RoboDK station: robotic_car_painting_cell.rdk

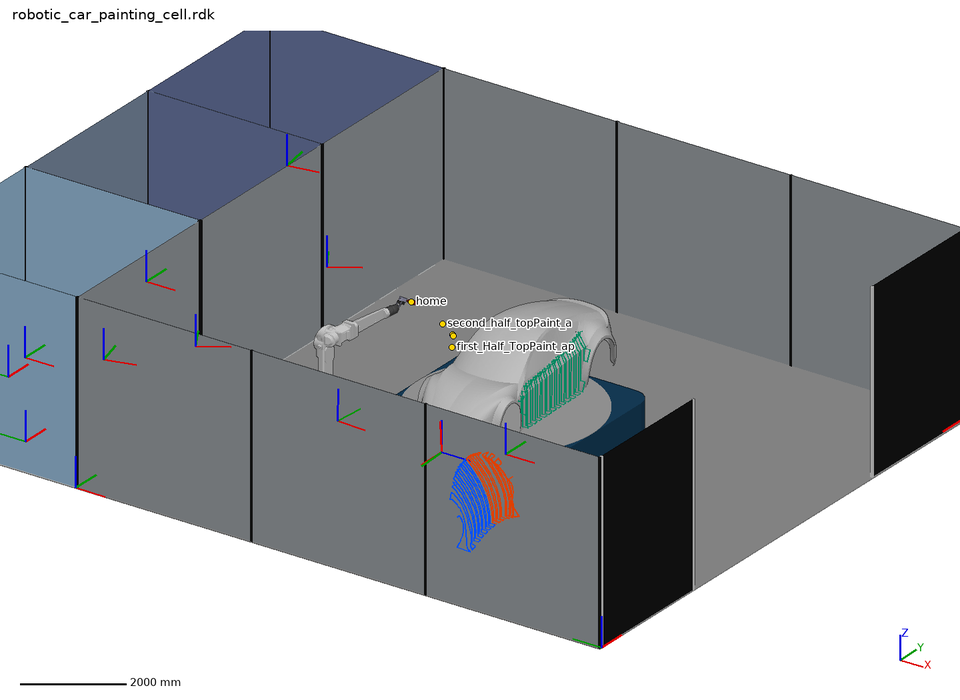
[picture v0: the station drawn from its stored meshes, robots at their saved joint values, targets as dots, program paths as lines]
Station robotic_car_painting_cell (saved by RoboDK 6.1.1). Poses are relative to the parent item; angles as X-Y-Z fixed-axis rotations.
  - frame ABB IRB 5500-27 Base at (-2375.69, -2107.7, 876.55) mm, rotated rx -0.57 ry -0.3 rz -4.19 deg
    - robot ABB IRB 5500-27: 6 axes, payload 16 kg, reach 2200 mm, repeatability 0.15 mm, weight 600 kg
        modified DH rows (alpha deg, a mm, theta deg, d mm): 0, 0, 0, 436; -90, 0, -90, -5; 0, 1300, 0, 0; -90, 0, -90, 1510.5; 35, 0, 0, 79.169; -70, 0, 180, 79.169
        base shift (0, 0, 0) mm, rotated rx 0 ry 0 rz 90 deg
        joint limits [-104, -65, -70, -719, -719, -720] to [104, 150, 70, 719, 719, 720]; home [0, 0, 0, 0, 0, 0]; saved at [0, 0, 0, 0, 0, 0]
      - tool Paint gun, TCP at (50, 0, 450) mm, rotated rx 0 ry 30 rz 0 deg, size 203.2 x 279.7 x 471.5 mm
    - target home (joint target) at (5, 2172.1, 1686) mm, rotated rx 180 ry 60 rz -90 deg; joints [0, 0, 0, 0, 0, 0, 0] of ABB IRB 5500-27
    - target first_Half_TopPaint_app (joint target) at (1861.11, 1119.96, 1686) mm, rotated rx 180 ry 60 rz -148.83 deg; joints [-58.83, 0, 0, 0, 0, 0, -69.91] of ABB IRB 5500-27
    - target second_half_topPaint_app (joint target) at (1072.69, 1796.81, 1679.78) mm, rotated rx 180 ry 59.9 rz -120.7 deg; joints [-30.7, -3.5, 3.6, 0, 0, 0, -28] of ABB IRB 5500-27
    - target second_to_home (joint target) at (1519.79, 1551.86, 1686) mm, rotated rx 180 ry 60 rz -134.27 deg; joints [-44.27, 0, 0, 0, 0, 0, -33.04] of ABB IRB 5500-27
    - target sidePaintApp (joint target) at (1560.69, 1510.73, 1686) mm, rotated rx 180 ry 60 rz -135.8 deg; joints [-45.8, 0, 0, 0, 0, 0, -170] of ABB IRB 5500-27
  - frame Turntable 1 Base at (0, 0, 0) mm
    - robot Turntable 1: 1 axes
        modified DH rows (alpha deg, a mm, theta deg, d mm): 0, 0, 0, 0
        base shift (0, 0, 1000) mm
        joint limits [-1000] to [1000]; home [0]; saved at [0]
      - frame carFrame at (0, -2099.21, -116.89) mm, rotated rx 90 ry 0 rz 0 deg
        - object carBodyTesla at (0, 0, 0) mm, size 1894.9 x 1628.8 x 4824.9 mm, geometry from carBodyTesla.STEP
        - frame FrameSidePaint at (0, 0, 0) mm, rotated rx -92.52 ry -89.99 rz 2.4 deg
          - object carSidePaint at (0, 0, 0) mm, geometry from       
        - frame FrameTopPaint at (0, 0, 0) mm, rotated rx 90 ry -3.48 rz 90 deg
          - object carTopPaint at (0, 0, 0) mm, rotated rx 90 ry 0 rz 86.52 deg, geometry from pacity
  - machining project first_half_topPaint: rotZ(0) | rotX(0)*rotY(0) | onStart | onPathStart | onApproach | onPoint | onRetract | onFinish | SetRPM(%1) | SetTool(%1) | Extruder(%1) | default | default | OutOnMov(%1) | OutOffMov(%1) | onPathFinish | M_RunCode(%1)
  - program first_half_topPaint (530 instructions, listed below)
  - machining project Path2 settings: rotZ(0) | rotX(0)*rotY(0) | rotz(0) | onStart | onPathStart | onApproach | onPoint | onRetract | onFinish | SetRPM(%1) | SetTool(%1) | Extruder(%1) | default | default | OutOnMov(%1) | OutOffMov(%1) | onPathFinish | M_RunCode(%1)
  - program second_half_topPaint (492 instructions, listed below)
  - machining project Path3 settings: rotZ(0) | rotX(0)*rotY(0) | rotz(90) | onStart | onPathStart | onApproach | onPoint | onRetract | onFinish | SetRPM(%1) | SetTool(%1) | Extruder(%1) | default | default | OutOnMov(%1) | OutOffMov(%1) | onPathFinish | M_RunCode(%1)
  - program side_paint (1096 instructions, listed below)
  - program second_half_topPaint_startP (3 instructions, listed below)
  - program first_half_topPaint_startP (3 instructions, listed below)
  - program second_to_First_conn (3 instructions, listed below)
  - program CarTopPaintMain (3 instructions, listed below)
  - program sidePaint_startP (3 instructions, listed below)
  - program CarSidePaintMain (1 instructions, listed below)
  - program Home (3 instructions, listed below)
  - object robot_stand at (-2371.87, -2116.55, 0) mm, size 1000 x 999.7 x 874.6 mm
  - frame Components at (-5797.63, -5825.6, 0) mm
    - frame Fence 1 Frame at (0, 0, 0) mm
      - object Fence 1 at (0, 0, 0) mm, size 12050 x 12050 x 4010 mm
    - frame Fence 1 Frame at (-4009.44, 0, 0) mm
      - object Fence 1 at (0, 0, 0) mm, size 4050 x 4050 x 4010 mm
    - frame Fence 1 Frame at (-3997.18, 4026.78, 0) mm
      - object Fence 1 at (0, 0, 0) mm, size 4050 x 4050 x 4010 mm
    - frame Fence 1 Frame at (-3995.72, 8010.06, 0) mm
      - object Fence 1 at (0, 0, 0) mm, size 4050 x 4050 x 4010 mm
    - frame Fence 1 Frame at (11995.78, 12001.82, 0) mm, rotated rx 0 ry 0 rz -90.05 deg
      - object Fence 1 at (0, 0, 0) mm, size 3050 x 50 x 4000 mm
    - frame Fence 2 Frame at (12049.84, 56.15, 0) mm, rotated rx 0 ry 0 rz 89.84 deg
      - object Fence 2 at (0, 0, 0) mm, size 3050 x 50 x 4000 mm
    - frame Box 1 Frame at (-1567.64, 10491.56, 0) mm, rotated rx 0 ry 0 rz 32.89 deg
      - object Box 1 at (0, 0, 0) mm, size 1000 x 1000 x 500 mm, geometry from cube.sld
    - frame Sphere 1 Frame at (-2358.15, 10303.8, 1975.89) mm, rotated rx 0 ry 0 rz 9.39 deg
      - object Sphere 1 at (0, -1304.1, -1382.72) mm, size 1000 x 1000 x 1000 mm, geometry from sph.sld
    - frame Prism 2 Frame at (-2731.49, 4804.46, 0) mm, rotated rx 0 ry 0 rz 14.89 deg
      - object Prism 2 at (0, 0, 0) mm, size 1000 x 1000 x 500 mm, geometry from prism.sld
    - frame Table 1 Frame at (-1857.36, 1009.43, 39.55) mm, rotated rx 0 ry 0 rz 90.42 deg
      - frame Table 1 Plane Frame at (-585.26, 0, 1600) mm
      - object Table 1 at (0, 0, 0) mm, size 2000 x 1000 x 1600 mm
    - frame Cone 1 Frame at (-1643.96, 6288.26, 0) mm, rotated rx 0 ry 0 rz 30.73 deg
      - object Cone 1 at (0, 0, 0) mm, size 700 x 700 x 600 mm
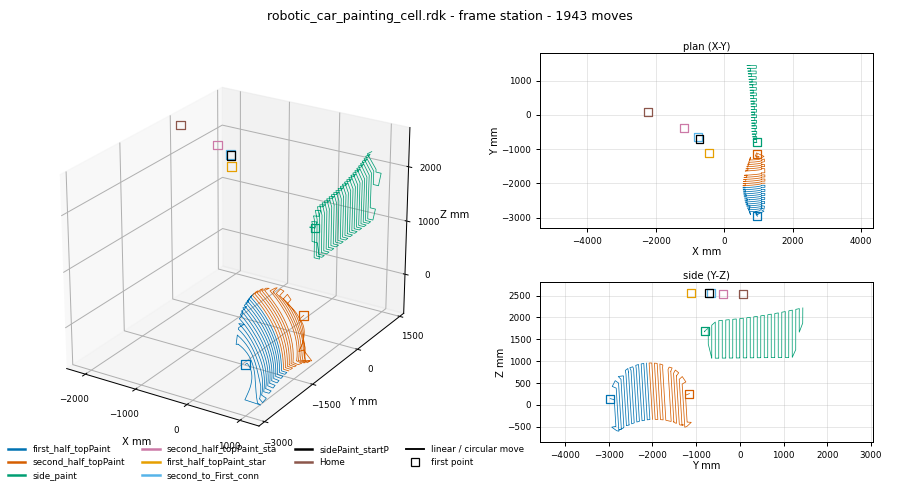
[picture p0: tool path of robotic_car_painting_cell.rdk in frame station, 1943 of 1943 moves have a stored position in this frame; points joined in program order, loops and branches not executed]

--- program first_half_topPaint (robot ABB IRB 5500-27) ---
  Smooth(1)
  Set speed (1000.0 mm/s)
  Set Ref.: FrameTopPaint
  Set Tool: Paint gun
  Show Paint gun
  MoveJ 1 to (-684.51, 907.52, 971.03) mm, rotated rx 106.25 ry 20.82 rz -12.55 deg; joints [-74.794, -12.721, 37.414, 15.51, -31.42, 69.743, -69.91]
  MoveL 2 to (-684.51, 907.52, 971.03) mm, rotated rx 106.25 ry 20.82 rz -12.55 deg; joints [-74.794, -12.721, 37.414, 15.51, -31.42, 69.743, -69.91]
  MoveL 3 to (-715.08, 815.97, 944.87) mm, rotated rx 106.25 ry 20.82 rz -12.55 deg; joints [-70.189, -11.053, 37.131, 20.085, -29.663, 64.32, -69.91]
  MoveL 4 to (-715.08, 815.97, 944.87) mm, rotated rx 106.25 ry 20.82 rz -12.55 deg; joints [-70.189, -11.053, 37.131, 20.085, -29.663, 64.32, -69.91]
  Set speed (50.0 mm/s)
  MoveL 5 to (-727.69, 815.97, 958.3) mm, rotated rx 115.21 ry 38.9 rz -3.5 deg; joints [-72.492, -7.954, 36.366, 53.545, -66.561, 43.021, -69.91]
  MoveL 6 to (-741.38, 815.97, 970.44) mm, rotated rx 121.28 ry 37.31 rz -1.34 deg; joints [-71.643, -9.484, 34.92, 41.962, -56.112, 42.571, -69.91]
  MoveL 7 to (-756.1, 815.97, 981.34) mm, rotated rx 127.91 ry 34.94 rz 0.84 deg; joints [-70.269, -10.891, 33.104, 25.851, -42.702, 44.586, -69.91]
  MoveL 8 to (-771.81, 815.97, 991.01) mm, rotated rx 147.14 ry 44.4 rz 22.43 deg; joints [-72.285, -8.078, 30.032, 38.203, -68.24, 34.256, -69.91]
  MoveL 9 to (-788.18, 815.97, 999.35) mm, rotated rx 152.65 ry 38.6 rz 23.9 deg; joints [-70.353, -9.282, 27.683, 18.408, -52.224, 37.943, -69.91]
  MoveL 10 to (-804.72, 815.97, 1006.28) mm, rotated rx 157.1 ry 32.58 rz 24.14 deg; joints [-67.802, -9.883, 25.248, -7.481, -33.792, 47.461, -69.91]
  MoveL 11 to (-821.7, 815.97, 1012.06) mm, rotated rx 171.62 ry 31.52 rz 45.71 deg; joints [-69.524, -6.36, 20.448, 5.697, -60.164, 39.026, -69.91]
  MoveL 12 to (-839.09, 815.97, 1016.77) mm, rotated rx 172.06 ry 25.49 rz 43.55 deg; joints [-67.355, -6.129, 18.073, -13.153, -47.594, 47.333, -69.91]
  MoveL 13 to (-856.8, 815.97, 1020.47) mm, rotated rx 172.25 ry 20.32 rz 41.61 deg; joints [-65.459, -5.39, 15.854, -31.628, -37.033, 57.574, -69.91]
  MoveL 14 to (-879.91, 815.97, 1023.85) mm, rotated rx 172.07 ry 15.06 rz 39.99 deg; joints [-63.836, -3.875, 13.191, -50.671, -28.335, 70.216, -69.91]
  MoveL 15 to (-903.07, 815.97, 1025.78) mm, rotated rx 171.26 ry 11.43 rz 39.86 deg; joints [-63.298, -1.925, 10.503, -57.68, -27.796, 76.89, -69.91]
  MoveL 16 to (-926.28, 815.97, 1026.44) mm, rotated rx 169.77 ry 9.41 rz 41.6 deg; joints [-63.721, 0.361, 7.673, -51.962, -34.901, 76.409, -69.91]
  MoveL 17 to (-949.54, 815.97, 1025.94) mm, rotated rx 167.69 ry 9.08 rz 45.24 deg; joints [-64.892, 2.979, 4.812, -39.109, -46.426, 72.324, -69.91]
  MoveL 18 to (-972.84, 815.97, 1024.4) mm, rotated rx 162.64 ry 4.98 rz 31.07 deg; joints [-63.067, 2.797, 5.746, -87.371, -13.884, 106.328, -69.91]
  MoveL 19 to (-996.1, 815.97, 1021.9) mm, rotated rx 159.46 ry 7.32 rz 37.29 deg; joints [-65.349, 5.612, 2.717, -48.527, -38.544, 85.33, -69.91]
  MoveL 20 to (-1019.16, 815.97, 1018.56) mm, rotated rx 156.28 ry 11.18 rz 43.19 deg; joints [-67.612, 8.569, 0.499, -24.443, -55.69, 75.354, -69.91]
  MoveL 21 to (-1054.91, 815.97, 1011.84) mm, rotated rx 147.55 ry 8.73 rz 32.21 deg; joints [-67.708, 9.55, 0.627, -38.437, -41.429, 89.233, -69.91]
  MoveL 22 to (-1090.21, 815.97, 1003.5) mm, rotated rx 141.46 ry 15.3 rz 35.63 deg; joints [-70.243, 13.119, -0.752, -11.462, -57.847, 79.186, -69.91]
  MoveL 23 to (-1125.14, 815.97, 993.72) mm, rotated rx 135.68 ry 21.23 rz 35.98 deg; joints [-71.841, 16.239, -1.381, 6.343, -68.344, 74.883, -69.91]
  MoveL 24 to (-1159.69, 815.96, 982.62) mm, rotated rx 130.17 ry 26.09 rz 34.38 deg; joints [-72.775, 18.955, -1.682, 19.317, -75.346, 72.813, -69.91]
  MoveL 25 to (-1193.94, 815.97, 970.3) mm, rotated rx 120.68 ry 12.99 rz 20.14 deg; joints [-71.511, 17.84, -0.657, -10.346, -46.92, 91.196, -69.91]
  MoveL 26 to (-1227.25, 815.97, 957.05) mm, rotated rx 116.07 ry 14.96 rz 18.47 deg; joints [-71.999, 19.907, -0.984, -1.213, -50.466, 88.745, -69.91]
  MoveL 27 to (-1260.2, 815.97, 942.74) mm, rotated rx 112.21 ry 16.36 rz 16.46 deg; joints [-72.228, 21.731, -1.288, 5.505, -52.512, 87.03, -69.91]
  MoveL 28 to (-1293.17, 815.97, 928.47) mm, rotated rx 109.24 ry 17.29 rz 14.07 deg; joints [-72.243, 23.194, -1.506, 9.979, -52.843, 85.592, -69.91]
  MoveL 29 to (-1326.13, 815.97, 914.18) mm, rotated rx 106.48 ry 18.02 rz 12.4 deg; joints [-72.245, 24.912, -2.196, 14.357, -54.013, 84.608, -69.91]
  Set speed (1000.0 mm/s)
  MoveL 30 to (-1326.13, 815.97, 914.18) mm, rotated rx 106.48 ry 18.02 rz 12.4 deg; joints [-72.245, 24.912, -2.196, 14.357, -54.013, 84.608, -69.91]
  MoveL 31 to (-1338.15, 911.5, 941.16) mm, rotated rx 106.48 ry 18.02 rz 12.4 deg; joints [-74.918, 25.452, -3.974, 14.165, -56.682, 86.948, -69.91]
  Set speed (1000.0 mm/s)
  MoveL 32 to (-1426.8, 802.28, 1164.66) mm, rotated rx 159.74 ry 21.34 rz 28.53 deg; joints [-65.232, 18.141, -13.203, -64.298, -13.867, 90.288, -69.91]
  MoveL 33 to (-1440.26, 755.54, 1077.29) mm, rotated rx 159.74 ry 21.34 rz 28.53 deg; joints [-63.808, 19.217, -11.228, -70.076, -7.316, 90.993, -69.91]
  MoveL 34 to (-1440.26, 755.54, 1077.29) mm, rotated rx 159.74 ry 21.34 rz 28.53 deg; joints [-63.808, 19.217, -11.228, -70.076, -7.316, 90.993, -69.91]
  Set speed (50.0 mm/s)
  MoveL 35 to (-1392.1, 755.54, 1069.69) mm, rotated rx 159.42 ry 21.04 rz 29.31 deg; joints [-64.03, 17.502, -9.102, -59.847, -13.964, 85.038, -69.91]
  MoveL 36 to (-1343.82, 755.54, 1063.71) mm, rotated rx 159.05 ry 20.67 rz 30.24 deg; joints [-64.278, 15.856, -7.078, -52.603, -19.082, 81.124, -69.91]
  MoveL 37 to (-1295.44, 755.54, 1059.53) mm, rotated rx 158.62 ry 20.22 rz 31.39 deg; joints [-64.567, 14.305, -5.248, -46.409, -23.965, 78.169, -69.91]
  MoveL 38 to (-1246.95, 755.54, 1056.8) mm, rotated rx 158.2 ry 19.77 rz 32.55 deg; joints [-64.842, 12.754, -3.469, -41.574, -28.141, 76.122, -69.91]
  MoveL 39 to (-1198.41, 755.54, 1054.98) mm, rotated rx 157.76 ry 19.27 rz 33.81 deg; joints [-65.127, 11.251, -1.802, -37.325, -32.182, 74.6, -69.91]
  MoveL 40 to (-1154.25, 755.54, 1053.79) mm, rotated rx 157.34 ry 18.77 rz 35.08 deg; joints [-65.394, 9.936, -0.387, -33.798, -35.852, 73.57, -69.91]
  MoveL 41 to (-1110.09, 755.54, 1052.74) mm, rotated rx 156.9 ry 18.21 rz 36.48 deg; joints [-65.67, 8.687, 0.922, -30.459, -39.626, 72.814, -69.91]
  MoveL 42 to (-1065.93, 755.54, 1051.53) mm, rotated rx 156.43 ry 17.58 rz 38.07 deg; joints [-65.958, 7.531, 2.102, -27.18, -43.642, 72.297, -69.91]
  MoveL 43 to (-1021.8, 755.54, 1049.88) mm, rotated rx 157.68 ry 19.17 rz 34.06 deg; joints [-65.149, 3.751, 6.657, -35.423, -33.05, 72.924, -69.91]
  MoveL 44 to (-977.72, 755.54, 1047.5) mm, rotated rx 167.62 ry 20.43 rz 49.37 deg; joints [-66.013, 3.469, 6.21, -13.59, -56.701, 56.758, -69.91]
  MoveL 45 to (-933.75, 755.54, 1044.07) mm, rotated rx 170.23 ry 16.63 rz 43.58 deg; joints [-63.285, -0.433, 9.362, -37.882, -37.374, 65.285, -69.91]
  MoveL 46 to (-889.98, 755.54, 1039.27) mm, rotated rx 173.11 ry 14.65 rz 38.16 deg; joints [-60.377, -4.093, 13.488, -83.022, -6.548, 88.314, -69.91]
  MoveL 47 to (-860.05, 755.54, 1035) mm, rotated rx -179.66 ry 15.22 rz 55.82 deg; joints [-62.992, -3.267, 11.61, -25.717, -52.157, 51.737, -69.91]
  MoveL 48 to (-830.27, 755.54, 1029.79) mm, rotated rx -177.87 ry 15.22 rz 53.67 deg; joints [-61.924, -5.683, 14.166, -32.954, -44.629, 52.598, -69.91]
  MoveL 49 to (-800.66, 755.54, 1023.53) mm, rotated rx -176.11 ry 16.07 rz 52.51 deg; joints [-61.237, -7.933, 16.745, -36.847, -39.487, 51.96, -69.91]
  MoveL 50 to (-771.23, 755.54, 1016.08) mm, rotated rx -174.42 ry 17.74 rz 52.38 deg; joints [-61.049, -10.014, 19.323, -35.956, -37.616, 48.908, -69.91]
  MoveL 51 to (-746.52, 755.54, 1008.72) mm, rotated rx -173.04 ry 19.78 rz 53.06 deg; joints [-61.359, -11.624, 21.506, -30.839, -39.113, 44.159, -69.91]
  MoveL 52 to (-722.23, 755.54, 1000.38) mm, rotated rx -171.69 ry 22.36 rz 54.42 deg; joints [-62.128, -13.046, 23.699, -22.211, -43.408, 37.945, -69.91]
  MoveL 53 to (-698.41, 755.54, 991.01) mm, rotated rx -170.31 ry 25.46 rz 56.4 deg; joints [-63.329, -14.226, 25.938, -11.163, -50.119, 31.19, -69.91]
  MoveL 54 to (-675.09, 755.54, 980.51) mm, rotated rx 179.52 ry 30.95 rz 35.88 deg; joints [-59.309, -18.43, 31.602, -48.712, -5.861, 51.566, -69.91]
  MoveL 55 to (-652.31, 755.54, 968.84) mm, rotated rx 179.13 ry 35.21 rz 37.82 deg; joints [-62.087, -19.133, 33.503, -8.823, -31.544, 29.317, -69.91]
  MoveL 56 to (-630.09, 755.54, 955.91) mm, rotated rx 178.55 ry 39.82 rz 39.79 deg; joints [-64.502, -19.381, 35.887, 12.39, -47.584, 20.25, -69.91]
  MoveL 57 to (-609.71, 755.54, 942.52) mm, rotated rx 159.64 ry 40.4 rz 14.9 deg; joints [-60.896, -22.487, 39.641, 4.355, -21.718, 26.226, -69.91]
  MoveL 58 to (-590.12, 755.54, 928.04) mm, rotated rx 155.96 ry 44.19 rz 14.66 deg; joints [-63.478, -22.211, 41.963, 27.837, -40.756, 17.955, -69.91]
  MoveL 59 to (-571.39, 755.54, 912.51) mm, rotated rx 151.85 ry 47.72 rz 13.83 deg; joints [-65.446, -21.467, 44.101, 43.056, -55.125, 15.532, -69.91]
  MoveL 60 to (-553.53, 755.54, 895.92) mm, rotated rx 147.33 ry 50.88 rz 12.41 deg; joints [-66.996, -20.317, 45.988, 55.196, -67.661, 15.527, -69.91]
  MoveL 61 to (-536.67, 755.54, 878.41) mm, rotated rx 127.47 ry 39.25 rz -10.05 deg; joints [-63.366, -23.419, 48.128, 49.258, -42.824, 20.834, -69.91]
  MoveL 62 to (-520.01, 755.54, 859.01) mm, rotated rx 122.75 ry 40.4 rz -11.27 deg; joints [-64.734, -22.221, 49.83, 59, -53.504, 21.747, -69.91]
  MoveL 63 to (-504.53, 755.54, 838.79) mm, rotated rx 118.45 ry 41.21 rz -12.44 deg; joints [-65.784, -20.803, 51.259, 66.816, -62.622, 23.506, -69.91]
  MoveL 64 to (-490.18, 755.54, 817.78) mm, rotated rx 114.61 ry 41.73 rz -13.49 deg; joints [-66.594, -19.238, 52.459, 73.414, -70.636, 25.633, -69.91]
  MoveL 65 to (-476.91, 755.54, 796.04) mm, rotated rx 106.99 ry 23.12 rz -22.12 deg; joints [-63.461, -23.239, 52.863, 50.56, -34.618, 37.619, -69.91]
  MoveL 66 to (-464.68, 755.54, 773.58) mm, rotated rx 104.59 ry 23.01 rz -21.81 deg; joints [-64.372, -21.966, 53.963, 56.36, -41.539, 38.387, -69.91]
  MoveL 67 to (-453.44, 755.54, 750.43) mm, rotated rx 102.53 ry 22.87 rz -21.47 deg; joints [-65.129, -20.575, 54.912, 61.159, -47.64, 39.407, -69.91]
  Set speed (1000.0 mm/s)
  MoveL 68 to (-453.44, 755.54, 750.43) mm, rotated rx 102.53 ry 22.87 rz -21.47 deg; joints [-65.129, -20.575, 54.912, 61.159, -47.64, 39.407, -69.91]
  MoveL 69 to (-409.87, 843.3, 770.43) mm, rotated rx 102.53 ry 22.87 rz -21.47 deg; joints [-71.111, -24.293, 56.106, 49.582, -44.096, 47.651, -69.91]
  Set speed (1000.0 mm/s)
  MoveL 70 to (-281.6, 768.08, 751.28) mm, rotated rx 118.7 ry 43.33 rz -18.27 deg; joints [-62.377, -34.976, 63.523, 74.349, -60.557, 13.693, -69.91]
  MoveL 71 to (-340.39, 695.12, 716.35) mm, rotated rx 118.7 ry 43.33 rz -18.27 deg; joints [-56.8, -27.468, 61.651, 88.642, -70.457, 7.211, -69.91]
  MoveL 72 to (-340.39, 695.12, 716.35) mm, rotated rx 118.7 ry 43.33 rz -18.27 deg; joints [-56.8, -27.468, 61.651, 88.642, -70.457, 7.211, -69.91]
  Set speed (50.0 mm/s)
  MoveL 73 to (-357.79, 695.12, 744.11) mm, rotated rx 122.68 ry 42.81 rz -17.25 deg; joints [-55.745, -29.267, 60.106, 82.857, -61.77, 3.52, -69.91]
  MoveL 74 to (-376.42, 695.12, 770.89) mm, rotated rx 126.99 ry 42.02 rz -16.17 deg; joints [-54.495, -30.632, 58.299, 76.918, -52.791, -0.116, -69.91]
  MoveL 75 to (-396.34, 695.12, 796.64) mm, rotated rx 148.49 ry 54.01 rz 7.6 deg; joints [-59.555, -28.01, 56.176, 69.276, -68.984, 0.456, -69.91]
  MoveL 76 to (-417.57, 695.12, 821.34) mm, rotated rx 153.05 ry 51.3 rz 9.14 deg; joints [-57.958, -29.273, 54.05, 59.05, -56.504, -1.277, -69.91]
  MoveL 77 to (-440.16, 695.12, 844.95) mm, rotated rx 157.24 ry 48.23 rz 10.14 deg; joints [-56.057, -29.952, 51.614, 47.146, -42.953, -1.501, -69.91]
  MoveL 78 to (-463.66, 695.12, 867.05) mm, rotated rx 160.94 ry 44.95 rz 10.58 deg; joints [-53.841, -30.026, 48.928, 31.405, -27.268, 1.327, -69.91]
  MoveL 79 to (-488.26, 695.12, 887.85) mm, rotated rx -177.23 ry 43.87 rz 37.69 deg; joints [-58.143, -27.481, 45.354, 19.418, -40.991, 6.249, -69.91]
  MoveL 80 to (-513.9, 695.12, 907.34) mm, rotated rx -176.74 ry 39.88 rz 35.84 deg; joints [-55.608, -27.028, 42.73, -3.171, -22.994, 15.838, -69.91]
  MoveL 81 to (-540.52, 695.12, 925.54) mm, rotated rx -162.84 ry 32.42 rz 57.85 deg; joints [-59.624, -23.369, 37.774, -0.094, -47.387, 14.917, -69.91]
  MoveL 82 to (-568.48, 695.12, 942.69) mm, rotated rx -164.33 ry 29.13 rz 55.28 deg; joints [-57.935, -22.308, 35.245, -15.197, -36.629, 22.96, -69.91]
  MoveL 83 to (-597.05, 695.12, 958.44) mm, rotated rx -165.72 ry 26.24 rz 53.18 deg; joints [-56.598, -20.945, 32.849, -31.04, -26.777, 32.675, -69.91]
  MoveL 84 to (-626.18, 695.12, 972.88) mm, rotated rx -167.06 ry 23.76 rz 51.59 deg; joints [-55.71, -19.364, 30.604, -46.953, -18.029, 43.399, -69.91]
  MoveL 85 to (-655.83, 695.11, 986.11) mm, rotated rx -168.39 ry 21.71 rz 50.56 deg; joints [-55.345, -17.631, 28.45, -60.642, -11.394, 53.406, -69.91]
  MoveL 86 to (-685.96, 695.11, 998.24) mm, rotated rx -169.75 ry 20.11 rz 50.1 deg; joints [-55.521, -15.787, 26.183, -65.849, -10.309, 58.613, -69.91]
  MoveL 87 to (-716.51, 695.11, 1009.37) mm, rotated rx -171.13 ry 18.97 rz 50.24 deg; joints [-56.138, -13.857, 23.731, -61.12, -15.403, 57.969, -69.91]
  MoveL 88 to (-747.45, 695.11, 1019.59) mm, rotated rx -172.55 ry 18.29 rz 50.98 deg; joints [-57.069, -11.851, 21.268, -52.76, -22.729, 55.229, -69.91]
  MoveL 89 to (-791.34, 695.11, 1032.58) mm, rotated rx 161.09 ry 5.65 rz 34.23 deg; joints [-59.026, -4.115, 12.605, -89.123, -11.867, 108.649, -69.91]
  MoveL 90 to (-835.67, 695.11, 1044.23) mm, rotated rx 160.86 ry 8.82 rz 33.33 deg; joints [-59.585, -3.228, 12.228, -94.03, -5.051, 109.893, -69.91]
  MoveL 91 to (-880.23, 695.11, 1054.81) mm, rotated rx -177.1 ry 15.23 rz 52.77 deg; joints [-59.128, -3.906, 11.744, -42.295, -36.545, 56.64, -69.91]
  MoveL 92 to (-924.96, 695.11, 1064.59) mm, rotated rx -176.34 ry 17.23 rz 53.99 deg; joints [-59.964, -2.248, 10.238, -35.087, -40.353, 51.827, -69.91]
  MoveL 93 to (-969.81, 695.11, 1073.86) mm, rotated rx -175.63 ry 18.97 rz 55.01 deg; joints [-60.663, -0.543, 8.653, -29.288, -43.512, 48.078, -69.91]
  MoveL 94 to (-1028.62, 695.11, 1085.64) mm, rotated rx -174.5 ry 21.13 rz 56.04 deg; joints [-61.373, 1.61, 6.639, -23.31, -46.499, 43.959, -69.91]
  MoveL 95 to (-1087.4, 695.11, 1097.53) mm, rotated rx -173.09 ry 23.15 rz 56.68 deg; joints [-61.836, 3.619, 4.728, -19.013, -48.087, 40.417, -69.91]
  MoveL 96 to (-1146.04, 695.11, 1110.05) mm, rotated rx 166.26 ry 15.84 rz 50.49 deg; joints [-63.474, 11.81, -6.483, -23.849, -54.817, 67.446, -69.91]
  MoveL 97 to (-1181.2, 695.11, 1109.5) mm, rotated rx 160.25 ry 10.46 rz 33.87 deg; joints [-61.223, 11.407, -5.811, -72.396, -19.793, 99.298, -69.91]
  MoveL 98 to (-1216.21, 695.11, 1107.75) mm, rotated rx 158.74 ry 10.98 rz 37.04 deg; joints [-62.275, 14.075, -9.07, -53.885, -32.649, 90.31, -69.91]
  MoveL 99 to (-1251.08, 695.11, 1104.82) mm, rotated rx 157.26 ry 11.78 rz 40.19 deg; joints [-63.246, 16.789, -12.164, -40.885, -42.47, 85.113, -69.91]
  MoveL 100 to (-1285.82, 695.11, 1100.76) mm, rotated rx 155.81 ry 12.84 rz 43.32 deg; joints [-64.127, 19.568, -15.232, -30.224, -51.075, 81.751, -69.91]
  MoveL 101 to (-1322.08, 695.11, 1095.31) mm, rotated rx 154.39 ry 14.16 rz 46.4 deg; joints [-64.923, 22.485, -18.398, -20.85, -58.987, 79.564, -69.91]
  MoveL 102 to (-1358.19, 695.11, 1088.66) mm, rotated rx 153.08 ry 15.63 rz 49.27 deg; joints [-65.598, 25.417, -21.571, -12.718, -66.093, 78.345, -69.91]
  MoveL 103 to (-1394.16, 695.11, 1080.85) mm, rotated rx 152.68 ry 16.63 rz 49.61 deg; joints [-65.828, 27.247, -23.476, -10.479, -67.345, 77.844, -69.91]
  Set speed (1000.0 mm/s)
  MoveL 104 to (-1394.16, 695.11, 1080.85) mm, rotated rx 152.68 ry 16.63 rz 49.61 deg; joints [-65.828, 27.247, -23.476, -10.479, -67.345, 77.844, -69.91]
  MoveL 105 to (-1412.65, 744.22, 1165.98) mm, rotated rx 152.68 ry 16.63 rz 49.61 deg; joints [-67.153, 27.921, -27.492, -9.895, -70.144, 81.333, -69.91]
  Set speed (1000.0 mm/s)
  MoveL 106 to (-1375.51, 652.07, 1179.39) mm, rotated rx 165.62 ry -5.87 rz 27.7 deg; joints [-57.069, 23.686, -26.713, -100.602, -28.973, 130.104, -69.91]
  MoveL 107 to (-1355.21, 634.69, 1083.02) mm, rotated rx 165.62 ry -5.87 rz 27.7 deg; joints [-56.558, 22.709, -21.583, -112.815, -18.302, 134.572, -69.91]
  MoveL 108 to (-1355.21, 634.69, 1083.02) mm, rotated rx 165.62 ry -5.87 rz 27.7 deg; joints [-56.558, 22.709, -21.583, -112.815, -18.302, 134.572, -69.91]
  Set speed (50.0 mm/s)
  MoveL 109 to (-1316.38, 634.69, 1090.54) mm, rotated rx 160.01 ry 2.28 rz 38.18 deg; joints [-59.418, 21.194, -19.149, -66.304, -35.59, 102.897, -69.91]
  MoveL 110 to (-1277.34, 634.69, 1096.75) mm, rotated rx 162.3 ry 1.08 rz 33.21 deg; joints [-58.086, 18.107, -15.194, -92.332, -19.797, 117.137, -69.91]
  MoveL 111 to (-1238.22, 634.69, 1101.6) mm, rotated rx 165.67 ry 5.56 rz 47.62 deg; joints [-59.572, 17.641, -15.337, -47.715, -46.895, 85.041, -69.91]
  MoveL 112 to (-1199.15, 634.69, 1105.05) mm, rotated rx 167.83 ry 4.65 rz 43.07 deg; joints [-58.188, 14.451, -11.494, -65.355, -34.029, 92.461, -69.91]
  MoveL 113 to (-1160.12, 634.69, 1107.1) mm, rotated rx 170.05 ry 4.26 rz 38.86 deg; joints [-56.822, 11.43, -7.504, -91.093, -17.145, 105.753, -69.91]
  MoveL 114 to (-1118.77, 634.69, 1107.71) mm, rotated rx 174.28 ry 6.72 rz 54.89 deg; joints [-58.543, 11.249, -8.209, -42.235, -50.513, 72.395, -69.91]
  MoveL 115 to (-1077.45, 634.69, 1106.69) mm, rotated rx 176.61 ry 6.55 rz 51.55 deg; joints [-57.243, 8.06, -4.378, -54.834, -39.766, 75.932, -69.91]
  MoveL 116 to (-1036.19, 634.69, 1104.01) mm, rotated rx 178.95 ry 6.82 rz 48.77 deg; joints [-55.954, 5.026, -0.567, -69.458, -28.178, 81.246, -69.91]
  MoveL 117 to (-994.97, 634.69, 1099.63) mm, rotated rx -178.75 ry 7.47 rz 46.55 deg; joints [-54.75, 2.128, 3.393, -91.116, -12.694, 91.284, -69.91]
  MoveL 118 to (-953.8, 634.69, 1093.51) mm, rotated rx -173.84 ry 6.74 rz 64.97 deg; joints [-57, 2.502, 1.816, -35.936, -55.36, 55.838, -69.91]
  MoveL 119 to (-912.68, 634.69, 1085.62) mm, rotated rx -172.59 ry 19.22 rz 52 deg; joints [-56.176, -4.46, 12.549, -52.051, -23.377, 55.8, -69.91]
  MoveL 120 to (-871.51, 634.69, 1072.56) mm, rotated rx -172.59 ry 19.22 rz 52 deg; joints [-55.881, -6.196, 14.647, -52.719, -22.54, 55.832, -69.91]
  MoveL 121 to (-830.42, 634.69, 1059.28) mm, rotated rx -172.59 ry 19.22 rz 52 deg; joints [-55.566, -7.94, 16.718, -53.538, -21.623, 55.98, -69.91]
  MoveL 122 to (-789.46, 634.69, 1045.61) mm, rotated rx -171.94 ry 19.13 rz 51.23 deg; joints [-54.643, -9.997, 19.236, -62.921, -14.618, 60.304, -69.91]
  MoveL 123 to (-748.7, 634.69, 1031.35) mm, rotated rx -156.77 ry 18 rz 70.54 deg; joints [-56.819, -11.685, 21.368, -19.559, -51.213, 24.851, -69.91]
  MoveL 124 to (-708.28, 634.69, 1016.36) mm, rotated rx -156.77 ry 18 rz 70.54 deg; joints [-56.513, -13.435, 23.355, -19.855, -50.662, 24.684, -69.91]
  MoveL 125 to (-668.3, 634.69, 1000.48) mm, rotated rx -156.77 ry 18 rz 70.54 deg; joints [-56.189, -15.177, 25.327, -20.186, -50.077, 24.537, -69.91]
  MoveL 126 to (-628.85, 634.69, 983.53) mm, rotated rx -156.77 ry 18 rz 70.54 deg; joints [-55.845, -16.906, 27.286, -20.548, -49.456, 24.401, -69.91]
  MoveL 127 to (-590.02, 634.69, 965.35) mm, rotated rx -156.77 ry 18 rz 70.54 deg; joints [-55.481, -18.618, 29.236, -20.935, -48.798, 24.266, -69.91]
  MoveL 128 to (-555.82, 634.69, 947.87) mm, rotated rx -156.77 ry 18 rz 70.54 deg; joints [-55.138, -20.133, 30.98, -21.295, -48.178, 24.134, -69.91]
  MoveL 129 to (-522.25, 634.69, 929.14) mm, rotated rx -154.84 ry 19.45 rz 71.77 deg; joints [-55.326, -21.996, 33.592, -16.618, -50.193, 19.687, -69.91]
  MoveL 130 to (-489.37, 634.69, 909.05) mm, rotated rx -152.75 ry 21.25 rz 73.54 deg; joints [-55.902, -23.696, 36.251, -9.884, -54.143, 14.522, -69.91]
  MoveL 131 to (-457.22, 634.69, 887.47) mm, rotated rx -160.07 ry 31.84 rz 55.32 deg; joints [-51.698, -28.268, 42.389, -19.018, -24.825, 16.788, -69.91]
  MoveL 132 to (-425.94, 634.69, 864.33) mm, rotated rx -158.53 ry 34.89 rz 57.9 deg; joints [-53.448, -29.496, 45.091, -0.084, -38.209, 6.341, -69.91]
  MoveL 133 to (-398.61, 634.69, 842.13) mm, rotated rx -173.74 ry 43.01 rz 35.04 deg; joints [-48.475, -32.48, 49.548, 9.522, -20.828, -0.175, -69.91]
  MoveL 134 to (-372.41, 634.69, 818.84) mm, rotated rx 165.27 ry 44.76 rz 8.05 deg; joints [-43.91, -33.935, 52.801, 50.133, -25.689, -21.91, -69.91]
  MoveL 135 to (-347.35, 634.69, 794.46) mm, rotated rx 162.46 ry 47.56 rz 7.96 deg; joints [-45.254, -34.584, 55.577, 59.853, -37.096, -22.308, -69.91]
  MoveL 136 to (-323.43, 634.69, 768.98) mm, rotated rx 159.27 ry 50.25 rz 7.51 deg; joints [-46.594, -34.742, 58.17, 67.86, -47.71, -21.078, -69.91]
  MoveL 137 to (-300.65, 634.69, 742.4) mm, rotated rx 155.72 ry 52.77 rz 6.66 deg; joints [-47.907, -34.337, 60.554, 75.272, -58.153, -18.915, -69.91]
  MoveL 138 to (-279, 634.7, 714.74) mm, rotated rx 151.82 ry 55.08 rz 5.38 deg; joints [-49.149, -33.306, 62.708, 82.622, -68.741, -16.078, -69.91]
  MoveL 139 to (-258.48, 634.69, 685.99) mm, rotated rx 129.3 ry 43.6 rz -19.78 deg; joints [-41.92, -34.474, 64.469, 105.319, -65.232, -20.768, -69.91]
  Set speed (1000.0 mm/s)
  MoveL 140 to (-258.48, 634.69, 685.99) mm, rotated rx 129.3 ry 43.6 rz -19.78 deg; joints [-41.92, -34.474, 64.469, 105.319, -65.232, -20.768, -69.91]
  MoveL 141 to (-191.18, 692.73, 731.86) mm, rotated rx 147.63 ry 57.11 rz 3.73 deg; joints [-54.053, -41.711, 66.692, 75.22, -66.189, -7.883, -69.91]
  Set speed (1000.0 mm/s)
  MoveL 142 to (-183.28, 575.62, 758.7) mm, rotated rx 177.1 ry 6.02 rz -19.07 deg; joints [-21.942, -26.066, 40.425, 184.05, -63.541, -117.802, -69.91]
  MoveL 143 to (-194.83, 574.27, 659.38) mm, rotated rx 177.1 ry 6.02 rz -19.07 deg; joints [-22.549, -24.032, 42.868, 178.777, -60.803, -112.433, -69.91]
  MoveL 144 to (-194.83, 574.27, 659.38) mm, rotated rx 177.1 ry 6.02 rz -19.07 deg; joints [-22.549, -24.032, 42.868, 178.777, -60.803, -112.433, -69.91]
  Set speed (50.0 mm/s)
  MoveL 145 to (-219.86, 574.27, 691.41) mm, rotated rx 177.1 ry 6.02 rz -19.07 deg; joints [-23.585, -23.551, 41.338, 178.027, -59.446, -113.685, -69.91]
  MoveL 146 to (-246.13, 574.27, 722.19) mm, rotated rx 177.1 ry 6.02 rz -19.07 deg; joints [-24.633, -22.958, 39.784, 177.203, -58.039, -114.83, -69.91]
  MoveL 147 to (-273.65, 574.26, 751.72) mm, rotated rx 177.1 ry 6.02 rz -19.07 deg; joints [-25.688, -22.261, 38.205, 176.313, -56.589, -115.871, -69.91]
  MoveL 148 to (-302.4, 574.26, 780.01) mm, rotated rx 177.1 ry 6.02 rz -19.07 deg; joints [-26.745, -21.468, 36.602, 175.363, -55.104, -116.814, -69.91]
  MoveL 149 to (-332.38, 574.26, 807.07) mm, rotated rx 177.1 ry 6.02 rz -19.07 deg; joints [-27.8, -20.585, 34.975, 174.359, -53.591, -117.665, -69.91]
  MoveL 150 to (-362.98, 574.26, 832.48) mm, rotated rx 177.1 ry 6.02 rz -19.07 deg; joints [-28.83, -19.637, 33.354, 173.331, -52.085, -118.415, -69.91]
  MoveL 151 to (-394.69, 574.26, 856.77) mm, rotated rx 177.1 ry 6.02 rz -19.07 deg; joints [-29.85, -18.615, 31.71, 172.266, -50.567, -119.088, -69.91]
  MoveL 152 to (-427.24, 574.26, 879.8) mm, rotated rx 177.1 ry 6.02 rz -19.07 deg; joints [-30.848, -17.533, 30.053, 171.182, -49.057, -119.685, -69.91]
  MoveL 153 to (-460.48, 574.26, 901.58) mm, rotated rx 177.1 ry 6.02 rz -19.07 deg; joints [-31.819, -16.4, 28.387, 170.091, -47.564, -120.214, -69.91]
  MoveL 154 to (-500.86, 574.26, 926.04) mm, rotated rx 177.1 ry 6.02 rz -19.07 deg; joints [-32.938, -14.992, 26.39, 168.794, -45.818, -120.768, -69.91]
  MoveL 155 to (-542.03, 574.26, 949.04) mm, rotated rx 177.1 ry 6.02 rz -19.07 deg; joints [-34.014, -13.53, 24.374, 167.515, -44.115, -121.257, -69.91]
  MoveL 156 to (-583.91, 574.26, 970.77) mm, rotated rx 177.1 ry 6.02 rz -19.07 deg; joints [-35.046, -12.021, 22.337, 166.27, -42.464, -121.699, -69.91]
  MoveL 157 to (-626.38, 574.26, 991.41) mm, rotated rx 177.1 ry 6.02 rz -19.07 deg; joints [-36.033, -10.472, 20.274, 165.077, -40.874, -122.111, -69.91]
  MoveL 158 to (-669.37, 574.26, 1011.13) mm, rotated rx 177.1 ry 6.02 rz -19.07 deg; joints [-36.973, -8.889, 18.181, 163.954, -39.354, -122.513, -69.91]
  MoveL 159 to (-712.75, 574.26, 1030.11) mm, rotated rx 177.1 ry 6.02 rz -19.07 deg; joints [-37.868, -7.278, 16.055, 162.922, -37.913, -122.925, -69.91]
  MoveL 160 to (-749.34, 574.26, 1044.06) mm, rotated rx 177.71 ry 6.27 rz -20.13 deg; joints [-38.082, -5.583, 14.069, 165.371, -40.265, -124.307, -69.91]
  MoveL 161 to (-786.23, 574.26, 1056.58) mm, rotated rx 177.71 ry 6.27 rz -20.13 deg; joints [-38.778, -4.189, 12.311, 164.55, -39.14, -124.597, -69.91]
  MoveL 162 to (-823.42, 574.26, 1067.67) mm, rotated rx 177.71 ry 6.27 rz -20.13 deg; joints [-39.448, -2.772, 10.553, 163.731, -38.041, -124.845, -69.91]
  MoveL 163 to (-860.92, 574.26, 1077.35) mm, rotated rx 177.71 ry 6.27 rz -20.13 deg; joints [-40.093, -1.33, 8.795, 162.913, -36.966, -125.055, -69.91]
  MoveL 164 to (-898.7, 574.26, 1085.6) mm, rotated rx -180 ry 0 rz -20 deg; joints [-41.182, 2.327, 3.58, 177.336, -40.791, -137.341, -69.91]
  MoveL 165 to (-936.11, 574.26, 1092.33) mm, rotated rx -180 ry 0 rz -20 deg; joints [-41.728, 3.806, 1.792, 177.063, -40.134, -137.806, -69.91]
  MoveL 166 to (-973.79, 574.26, 1097.7) mm, rotated rx -180 ry 0 rz -20 deg; joints [-42.256, 5.308, -0.004, 176.796, -39.496, -138.247, -69.91]
  MoveL 167 to (-1011.76, 574.26, 1101.72) mm, rotated rx -180 ry 0 rz -20 deg; joints [-42.765, 6.834, -1.81, 176.537, -38.877, -138.667, -69.91]
  MoveL 168 to (-1050.02, 574.26, 1104.38) mm, rotated rx -180 ry 0 rz -20 deg; joints [-43.257, 8.385, -3.627, 176.286, -38.279, -139.067, -69.91]
  MoveL 169 to (-1095.85, 574.26, 1105.77) mm, rotated rx -180 ry 0 rz -20 deg; joints [-43.82, 10.263, -5.806, 175.999, -37.593, -139.522, -69.91]
  MoveL 170 to (-1141.59, 574.26, 1105.24) mm, rotated rx -180 ry 0 rz -20 deg; joints [-44.355, 12.157, -7.985, 175.732, -36.942, -139.954, -69.91]
  MoveL 171 to (-1187.18, 574.26, 1102.86) mm, rotated rx -180 ry 0 rz -20 deg; joints [-44.864, 14.069, -10.168, 175.487, -36.328, -140.366, -69.91]
  MoveL 172 to (-1232.62, 574.26, 1098.66) mm, rotated rx -180 ry 0 rz -20 deg; joints [-45.347, 15.999, -12.358, 175.267, -35.75, -140.764, -69.91]
  MoveL 173 to (-1277.91, 574.26, 1092.68) mm, rotated rx -180 ry 0 rz -20 deg; joints [-45.807, 17.95, -14.561, 175.075, -35.208, -141.154, -69.91]
  MoveL 174 to (-1323.07, 574.26, 1084.97) mm, rotated rx -180 ry 0 rz -20 deg; joints [-46.244, 19.924, -16.782, 174.917, -34.705, -141.541, -69.91]
  Set speed (1000.0 mm/s)
  MoveL 175 to (-1323.07, 574.26, 1084.97) mm, rotated rx -180 ry 0 rz -20 deg; joints [-46.244, 19.924, -16.782, 174.917, -34.705, -141.541, -69.91]
  MoveL 176 to (-1323.07, 574.26, 1184.97) mm, rotated rx -180 ry 0 rz -20 deg; joints [-46.083, 19.935, -20.429, 183.463, -39.574, -147.955, -69.91]
  Set speed (1000.0 mm/s)
  MoveL 177 to (-1313.47, 509.8, 1185.18) mm, rotated rx -176.65 ry -9.39 rz -6.29 deg; joints [-45.851, 23.319, -26.453, 203.524, -38.882, -173.412, -69.91]
  MoveL 178 to (-1296.65, 513.83, 1086.68) mm, rotated rx -176.65 ry -9.39 rz -6.29 deg; joints [-46.006, 22.269, -21.38, 192.12, -31.141, -166.393, -69.91]
  MoveL 179 to (-1296.65, 513.83, 1086.68) mm, rotated rx -176.65 ry -9.39 rz -6.29 deg; joints [-46.006, 22.269, -21.38, 192.12, -31.141, -166.393, -69.91]
  Set speed (50.0 mm/s)
  MoveL 180 to (-1253.37, 513.83, 1093.31) mm, rotated rx -177.02 ry -7.45 rz -5.52 deg; joints [-45.753, 19.397, -17.613, 181.453, -24.532, -160.148, -69.91]
  MoveL 181 to (-1210.06, 513.83, 1098.38) mm, rotated rx -177.41 ry -5.46 rz -4.72 deg; joints [-45.582, 16.581, -14.013, 167.425, -16.213, -151.616, -69.91]
  MoveL 182 to (-1166.74, 513.83, 1101.88) mm, rotated rx -176.77 ry -2.49 rz -23.92 deg; joints [-41.997, 16.522, -13.615, 193.52, -52.956, -147.223, -69.91]
  MoveL 183 to (-1123.4, 513.83, 1103.8) mm, rotated rx -177.87 ry -0.69 rz -23.09 deg; joints [-41.512, 13.747, -9.978, 187.882, -49.679, -143.405, -69.91]
  MoveL 184 to (-1080.04, 513.83, 1104.09) mm, rotated rx -179.01 ry 1.15 rz -22.28 deg; joints [-41.021, 11.014, -6.421, 182.051, -46.507, -139.289, -69.91]
  MoveL 185 to (-1036.65, 513.83, 1102.75) mm, rotated rx 179.82 ry 3.02 rz -21.49 deg; joints [-40.521, 8.316, -2.931, 176.025, -43.454, -134.863, -69.91]
  MoveL 186 to (-993.25, 513.83, 1099.72) mm, rotated rx 178.62 ry 4.93 rz -20.73 deg; joints [-40.01, 5.653, 0.497, 169.848, -40.563, -130.143, -69.91]
  MoveL 187 to (-949.82, 513.83, 1094.98) mm, rotated rx 177.38 ry 6.89 rz -20 deg; joints [-39.484, 3.019, 3.874, 163.569, -37.877, -125.148, -69.91]
  MoveL 188 to (-910.92, 513.83, 1089.24) mm, rotated rx 176.23 ry 8.67 rz -19.38 deg; joints [-38.995, 0.685, 6.861, 157.928, -35.693, -120.479, -69.91]
  MoveL 189 to (-872.4, 513.83, 1082.14) mm, rotated rx 175.05 ry 10.46 rz -18.81 deg; joints [-38.489, -1.605, 9.791, 152.415, -33.796, -115.72, -69.91]
  MoveL 190 to (-834.35, 513.83, 1073.7) mm, rotated rx 175.05 ry 10.46 rz -18.81 deg; joints [-37.782, -3.045, 11.508, 153.763, -35.202, -115.85, -69.91]
  MoveL 191 to (-796.77, 513.83, 1063.95) mm, rotated rx 175.05 ry 10.46 rz -18.81 deg; joints [-37.051, -4.454, 13.214, 155.094, -36.622, -115.931, -69.91]
  MoveL 192 to (-759.66, 513.83, 1052.88) mm, rotated rx 175.05 ry 10.46 rz -18.81 deg; joints [-36.295, -5.833, 14.91, 156.409, -38.058, -115.961, -69.91]
  MoveL 193 to (-720.8, 513.83, 1039.73) mm, rotated rx 175.05 ry 10.46 rz -18.81 deg; joints [-35.466, -7.261, 16.7, 157.79, -39.602, -115.937, -69.91]
  MoveL 194 to (-682.45, 513.83, 1025.14) mm, rotated rx 175.05 ry 10.46 rz -18.81 deg; joints [-34.605, -8.654, 18.481, 159.161, -41.17, -115.855, -69.91]
  MoveL 195 to (-644.6, 513.83, 1009.13) mm, rotated rx 175.05 ry 10.46 rz -18.81 deg; joints [-33.714, -10.011, 20.255, 160.526, -42.765, -115.712, -69.91]
  MoveL 196 to (-607.25, 513.83, 991.72) mm, rotated rx 175.05 ry 10.46 rz -18.81 deg; joints [-32.789, -11.33, 22.023, 161.888, -44.389, -115.509, -69.91]
  MoveL 197 to (-570.39, 513.83, 972.93) mm, rotated rx 175.05 ry 10.46 rz -18.81 deg; joints [-31.83, -12.611, 23.785, 163.252, -46.046, -115.244, -69.91]
  MoveL 198 to (-534.01, 513.83, 952.79) mm, rotated rx 175.05 ry 10.46 rz -18.81 deg; joints [-30.836, -13.852, 25.542, 164.623, -47.738, -114.915, -69.91]
  MoveL 199 to (-495.18, 513.83, 930.63) mm, rotated rx 175.05 ry 10.46 rz -18.81 deg; joints [-29.717, -15.159, 27.403, 166.167, -49.627, -114.545, -69.91]
  MoveL 200 to (-456.89, 513.83, 907.57) mm, rotated rx 175.05 ry 10.46 rz -18.81 deg; joints [-28.553, -16.422, 29.241, 167.752, -51.571, -114.128, -69.91]
  MoveL 201 to (-419.22, 513.83, 883.5) mm, rotated rx 175.05 ry 10.46 rz -18.81 deg; joints [-27.344, -17.634, 31.055, 169.369, -53.564, -113.65, -69.91]
  MoveL 202 to (-382.39, 513.83, 858.41) mm, rotated rx 175.05 ry 10.46 rz -18.81 deg; joints [-26.098, -18.783, 32.842, 171, -55.593, -113.099, -69.91]
  MoveL 203 to (-346.52, 513.84, 832.24) mm, rotated rx 175.05 ry 10.46 rz -18.81 deg; joints [-24.82, -19.862, 34.6, 172.637, -57.648, -112.467, -69.91]
  MoveL 204 to (-314.79, 513.84, 807.46) mm, rotated rx 175.05 ry 10.46 rz -18.81 deg; joints [-23.633, -20.774, 36.173, 174.121, -59.532, -111.812, -69.91]
  MoveL 205 to (-283.94, 513.84, 781.68) mm, rotated rx 175.05 ry 10.46 rz -18.81 deg; joints [-22.426, -21.614, 37.725, 175.596, -61.424, -111.073, -69.91]
  MoveL 206 to (-254.01, 513.84, 754.86) mm, rotated rx 178.74 ry 14.95 rz 1.79 deg; joints [-26.687, -27.559, 42.502, 104.602, -11.167, -87.381, -69.91]
  MoveL 207 to (-225.04, 513.84, 726.96) mm, rotated rx 178.61 ry 16.94 rz 1.9 deg; joints [-24.865, -28.845, 45.136, 114.092, -20.336, -90.65, -69.91]
  MoveL 208 to (-197.04, 513.84, 697.96) mm, rotated rx 178.48 ry 18.94 rz 2 deg; joints [-22.974, -29.966, 47.625, 120.393, -27.65, -91.844, -69.91]
  MoveL 209 to (-170.05, 513.84, 667.83) mm, rotated rx 178.29 ry 21.94 rz 2.11 deg; joints [-20.727, -31.055, 50.433, 126.011, -35.964, -91.718, -69.91]
  MoveL 210 to (-144.08, 513.84, 636.54) mm, rotated rx -138.81 ry 41.51 rz 59.54 deg; joints [-27.865, -37.22, 63.772, 56.737, -44.542, -59.045, -69.91]
  Set speed (1000.0 mm/s)
  MoveL 211 to (-144.08, 513.84, 636.54) mm, rotated rx -138.81 ry 41.51 rz 59.54 deg; joints [-27.865, -37.22, 63.772, 56.737, -44.542, -59.045, -69.91]
  MoveL 212 to (-62.03, 523.44, 692.89) mm, rotated rx -138.81 ry 41.51 rz 59.54 deg; joints [-22.624, -46.058, 64.763, 42.217, -26.661, -56.461, -69.91]
  Set speed (1000.0 mm/s)
  MoveL 213 to (-21.33, 463.02, 673.84) mm, rotated rx -138.81 ry 41.51 rz 59.54 deg; joints [-16.212, -43.404, 64.907, 61.194, -34.933, -69.907, -69.91]
  MoveL 214 to (-103.38, 453.41, 617.49) mm, rotated rx -138.81 ry 41.51 rz 59.54 deg; joints [-21.547, -35.141, 63.912, 68.724, -48.614, -67.825, -69.91]
  MoveL 215 to (-103.38, 453.41, 617.49) mm, rotated rx -138.81 ry 41.51 rz 59.54 deg; joints [-21.547, -35.141, 63.912, 68.724, -48.614, -67.825, -69.91]
  Set speed (50.0 mm/s)
  MoveL 216 to (-129.96, 453.41, 648.05) mm, rotated rx -140.91 ry 40.29 rz 58.16 deg; joints [-23.104, -35.66, 61.816, 58.446, -40.129, -62.315, -69.91]
  MoveL 217 to (-157.43, 453.41, 677.62) mm, rotated rx -160.08 ry 48.76 rz 32.41 deg; joints [-17.829, -31.302, 60.487, 107.365, -64.598, -76.049, -69.91]
  MoveL 218 to (-185.77, 453.41, 706.23) mm, rotated rx -161.37 ry 46.96 rz 31.44 deg; joints [-19.817, -31.67, 58.466, 99.981, -56.455, -74.357, -69.91]
  MoveL 219 to (-214.96, 453.41, 733.9) mm, rotated rx -162.58 ry 45.14 rz 30.55 deg; joints [-21.71, -31.683, 56.326, 92.184, -48.412, -71.875, -69.91]
  MoveL 220 to (-244.97, 453.41, 760.65) mm, rotated rx 176.48 ry 45.59 rz 1.76 deg; joints [-16.476, -27.043, 53.322, 137.489, -74.353, -79.89, -69.91]
  MoveL 221 to (-275.2, 453.41, 786.08) mm, rotated rx 176.68 ry 43.6 rz 1.88 deg; joints [-18.458, -26.862, 51.303, 132.518, -67.417, -80.649, -69.91]
  MoveL 222 to (-306.16, 453.41, 810.71) mm, rotated rx 176.87 ry 41.6 rz 1.98 deg; joints [-20.374, -26.444, 49.195, 127.622, -60.678, -81.042, -69.91]
  MoveL 223 to (-337.8, 453.41, 834.58) mm, rotated rx 177.05 ry 39.61 rz 2.06 deg; joints [-22.218, -25.819, 47.005, 122.686, -54.054, -81.081, -69.91]
  MoveL 224 to (-370.09, 453.41, 857.74) mm, rotated rx 177.22 ry 37.61 rz 2.12 deg; joints [-23.987, -25.012, 44.735, 117.581, -47.455, -80.745, -69.91]
  MoveL 225 to (-405.27, 453.41, 882.85) mm, rotated rx 177.37 ry 35.62 rz 2.17 deg; joints [-25.772, -23.999, 42.246, 111.834, -40.505, -79.898, -69.91]
  MoveL 226 to (-441.01, 453.41, 906.88) mm, rotated rx 177.52 ry 33.62 rz 2.21 deg; joints [-27.459, -22.829, 39.675, 105.414, -33.28, -78.42, -69.91]
  MoveL 227 to (-477.35, 453.41, 929.77) mm, rotated rx 177.66 ry 31.62 rz 2.23 deg; joints [-29.046, -21.519, 37.01, 97.672, -25.385, -75.95, -69.91]
  MoveL 228 to (-514.32, 453.41, 951.42) mm, rotated rx 177.8 ry 29.63 rz 2.23 deg; joints [-30.51, -20.08, 34.198, 86.701, -15.648, -71.354, -69.91]
  MoveL 229 to (-551.95, 453.41, 971.81) mm, rotated rx 166.35 ry 24.34 rz -17.72 deg; joints [-28.515, -16.34, 30.864, 144.542, -49.035, -92.27, -69.91]
  MoveL 230 to (-590.26, 453.41, 990.88) mm, rotated rx 167.62 ry 22.7 rz -17.83 deg; joints [-29.613, -14.53, 28.166, 145.007, -46.832, -95.01, -69.91]
  MoveL 231 to (-629.28, 453.41, 1008.58) mm, rotated rx 168.84 ry 21.04 rz -17.98 deg; joints [-30.671, -12.648, 25.435, 145.823, -44.905, -97.851, -69.91]
  MoveL 232 to (-665.67, 453.41, 1023.59) mm, rotated rx 170.01 ry 19.4 rz -18.16 deg; joints [-31.598, -10.818, 22.831, 147.168, -43.465, -100.804, -69.91]
  MoveL 233 to (-702.69, 453.41, 1037.4) mm, rotated rx 171.19 ry 17.67 rz -18.39 deg; joints [-32.483, -8.899, 20.152, 149.089, -42.409, -104.044, -69.91]
  MoveL 234 to (-740.35, 453.41, 1049.99) mm, rotated rx 172.34 ry 15.92 rz -18.67 deg; joints [-33.329, -6.909, 17.421, 151.501, -41.744, -107.479, -69.91]
  MoveL 235 to (-778.44, 453.41, 1061.25) mm, rotated rx 173.47 ry 14.16 rz -18.99 deg; joints [-34.134, -4.863, 14.653, 154.359, -41.47, -111.066, -69.91]
  MoveL 236 to (-816.69, 453.41, 1071.13) mm, rotated rx 174.56 ry 12.4 rz -19.34 deg; joints [-34.898, -2.777, 11.865, 157.61, -41.578, -114.758, -69.91]
  MoveL 237 to (-855.09, 453.41, 1079.64) mm, rotated rx 175.62 ry 10.65 rz -19.73 deg; joints [-35.623, -0.654, 9.05, 161.205, -42.042, -118.525, -69.91]
  MoveL 238 to (-901.38, 453.41, 1088.06) mm, rotated rx 176.85 ry 8.57 rz -20.22 deg; joints [-36.449, 1.941, 5.631, 165.885, -43.023, -123.094, -69.91]
  MoveL 239 to (-947.9, 453.41, 1094.56) mm, rotated rx 178.03 ry 6.5 rz -20.74 deg; joints [-37.235, 4.583, 2.163, 170.846, -44.398, -127.644, -69.91]
  MoveL 240 to (-994.63, 453.41, 1099.15) mm, rotated rx 179.16 ry 4.45 rz -21.28 deg; joints [-37.988, 7.274, -1.365, 175.996, -46.109, -132.127, -69.91]
  MoveL 241 to (-1041.57, 453.41, 1101.86) mm, rotated rx -179.75 ry 2.43 rz -21.82 deg; joints [-38.713, 10.016, -4.964, 181.259, -48.101, -136.503, -69.91]
  MoveL 242 to (-1088.73, 453.41, 1102.7) mm, rotated rx -178.7 ry 0.41 rz -22.35 deg; joints [-39.417, 12.808, -8.642, 186.555, -50.31, -140.736, -69.91]
  MoveL 243 to (-1135.25, 453.41, 1101.71) mm, rotated rx -177.72 ry -1.55 rz -22.85 deg; joints [-40.093, 15.605, -12.343, 191.746, -52.648, -144.742, -69.91]
  MoveL 244 to (-1181.97, 453.41, 1098.94) mm, rotated rx -178.19 ry -4.38 rz -3.27 deg; joints [-44.049, 15.682, -12.868, 158.004, -10.899, -145.001, -69.91]
  MoveL 245 to (-1228.61, 453.41, 1094.42) mm, rotated rx -178.04 ry -6.49 rz -3.6 deg; joints [-44.356, 18.557, -16.488, 174.541, -19.821, -155.599, -69.91]
  MoveL 246 to (-1275.06, 453.41, 1088.18) mm, rotated rx -177.96 ry -8.56 rz -3.79 deg; joints [-44.766, 21.471, -20.292, 186.498, -26.219, -163.227, -69.91]
  Set speed (1000.0 mm/s)
  MoveL 247 to (-1275.06, 453.41, 1088.18) mm, rotated rx -177.96 ry -8.56 rz -3.79 deg; joints [-44.766, 21.471, -20.292, 186.498, -26.219, -163.227, -69.91]
  MoveL 248 to (-1290.14, 450.85, 1187.01) mm, rotated rx -177.96 ry -8.56 rz -3.79 deg; joints [-44.603, 22.38, -25.162, 199.372, -34.626, -171.268, -69.91]
  Set speed (1000.0 mm/s)
  MoveL 249 to (-1271.01, 391.49, 1188.57) mm, rotated rx -178.86 ry -7.65 rz -2.1 deg; joints [-43.218, 21.855, -24.397, 195.392, -31.576, -168.653, -69.91]
  MoveL 250 to (-1257.64, 392.98, 1089.47) mm, rotated rx -178.86 ry -7.65 rz -2.1 deg; joints [-43.395, 21.066, -19.705, 181.218, -22.597, -159.678, -69.91]
  MoveL 251 to (-1257.64, 392.98, 1089.47) mm, rotated rx -178.86 ry -7.65 rz -2.1 deg; joints [-43.395, 21.066, -19.705, 181.218, -22.597, -159.678, -69.91]
  Set speed (50.0 mm/s)
  MoveL 252 to (-1213.67, 392.98, 1094.68) mm, rotated rx -178.71 ry -5.75 rz -2.36 deg; joints [-42.879, 18.442, -16.284, 170.271, -17.478, -152.253, -69.91]
  MoveL 253 to (-1169.62, 392.98, 1098.4) mm, rotated rx -178.64 ry -3.81 rz -2.43 deg; joints [-42.429, 15.852, -13.01, 156.276, -10.633, -142.88, -69.91]
  MoveL 254 to (-1125.48, 392.98, 1100.62) mm, rotated rx -178.11 ry -1.27 rz -22.37 deg; joints [-38.392, 16.135, -12.938, 192.598, -54.192, -143.869, -69.91]
  MoveL 255 to (-1081.26, 392.98, 1101.32) mm, rotated rx -178.86 ry 0.58 rz -22.19 deg; joints [-37.63, 13.614, -9.55, 188.452, -52.862, -140.274, -69.91]
  MoveL 256 to (-1036.98, 392.98, 1100.44) mm, rotated rx -179.68 ry 2.45 rz -21.95 deg; joints [-36.845, 11.124, -6.214, 184.357, -51.662, -136.618, -69.91]
  MoveL 257 to (-990.3, 392.98, 1097.8) mm, rotated rx 179.41 ry 4.44 rz -21.65 deg; joints [-35.987, 8.535, -2.748, 180.132, -50.583, -132.705, -69.91]
  MoveL 258 to (-943.96, 392.98, 1093.38) mm, rotated rx 178.44 ry 6.43 rz -21.33 deg; joints [-35.099, 6.003, 0.646, 176.095, -49.758, -128.782, -69.91]
  MoveL 259 to (-897.95, 392.98, 1087.19) mm, rotated rx 177.43 ry 8.42 rz -20.99 deg; joints [-34.175, 3.527, 3.976, 172.298, -49.231, -124.87, -69.91]
  MoveL 260 to (-852.29, 392.98, 1079.23) mm, rotated rx 176.38 ry 10.42 rz -20.66 deg; joints [-33.209, 1.107, 7.25, 168.796, -49.04, -120.994, -69.91]
  MoveL 261 to (-806.98, 392.98, 1069.48) mm, rotated rx 175.28 ry 12.42 rz -20.34 deg; joints [-32.195, -1.255, 10.474, 165.648, -49.224, -117.183, -69.91]
  MoveL 262 to (-762, 392.98, 1057.93) mm, rotated rx 174.15 ry 14.43 rz -20.05 deg; joints [-31.126, -3.553, 13.652, 162.915, -49.817, -113.469, -69.91]
  MoveL 263 to (-717.38, 392.98, 1044.57) mm, rotated rx 172.97 ry 16.43 rz -19.79 deg; joints [-29.997, -5.785, 16.789, 160.634, -50.839, -109.869, -69.91]
  MoveL 264 to (-673.11, 392.98, 1029.38) mm, rotated rx 171.74 ry 18.43 rz -19.57 deg; joints [-28.801, -7.945, 19.889, 158.835, -52.304, -106.394, -69.91]
  MoveL 265 to (-629.35, 392.98, 1012.43) mm, rotated rx 170.48 ry 20.4 rz -19.4 deg; joints [-27.538, -10.017, 22.939, 157.552, -54.211, -103.069, -69.91]
  MoveL 266 to (-586.54, 392.98, 993.9) mm, rotated rx 169.2 ry 22.34 rz -19.28 deg; joints [-26.215, -11.973, 25.91, 156.798, -56.533, -99.923, -69.91]
  MoveL 267 to (-544.68, 392.98, 973.85) mm, rotated rx 177.47 ry 26.8 rz 2.77 deg; joints [-29.633, -17.158, 29.972, 75.927, -5.018, -66.628, -69.91]
  MoveL 268 to (-503.74, 392.98, 952.35) mm, rotated rx 177 ry 28.93 rz 3.1 deg; joints [-28.409, -18.946, 33.24, 91.171, -17.641, -73.5, -69.91]
  MoveL 269 to (-460.08, 392.98, 927.29) mm, rotated rx 176.48 ry 30.82 rz 3.45 deg; joints [-26.991, -20.729, 36.305, 98.445, -25.083, -75.599, -69.91]
  MoveL 270 to (-417.43, 392.98, 900.62) mm, rotated rx 176.02 ry 31.78 rz 3.78 deg; joints [-25.616, -22.304, 38.862, 103.039, -29.699, -76.686, -69.91]
  MoveL 271 to (-375.74, 392.98, 872.42) mm, rotated rx 175.54 ry 32.73 rz 4.1 deg; joints [-24.173, -23.786, 41.374, 107.18, -34.106, -77.387, -69.91]
  MoveL 272 to (-334.95, 392.98, 842.8) mm, rotated rx 175.05 ry 33.68 rz 4.42 deg; joints [-22.659, -25.167, 43.844, 111.054, -38.421, -77.799, -69.91]
  MoveL 273 to (-294.98, 392.98, 811.84) mm, rotated rx 174.52 ry 34.62 rz 4.72 deg; joints [-21.069, -26.441, 46.274, 114.776, -42.72, -77.976, -69.91]
  MoveL 274 to (-255.76, 392.98, 779.72) mm, rotated rx 173.98 ry 35.56 rz 5.02 deg; joints [-19.393, -27.597, 48.662, 118.433, -47.059, -77.953, -69.91]
  MoveL 275 to (-217.15, 392.98, 746.61) mm, rotated rx 173.41 ry 36.49 rz 5.31 deg; joints [-17.622, -28.627, 51.006, 122.092, -51.482, -77.749, -69.91]
  MoveL 276 to (-217.15, 392.98, 746.61) mm, rotated rx 172.81 ry 37.42 rz 5.58 deg; joints [-17.913, -28.885, 51.487, 120.69, -51.803, -76.028, -69.91]
  MoveL 277 to (-183.3, 392.98, 716.57) mm, rotated rx 172.19 ry 38.33 rz 5.84 deg; joints [-16.3, -29.707, 53.579, 123.892, -55.891, -75.548, -69.91]
  MoveL 278 to (-150.38, 392.98, 685.6) mm, rotated rx 171.55 ry 39.24 rz 6.08 deg; joints [-14.63, -30.368, 55.624, 127.144, -60.108, -74.881, -69.91]
  MoveL 279 to (-123.21, 392.98, 658.55) mm, rotated rx 171.3 ry 40.23 rz 5.97 deg; joints [-12.715, -30.478, 57.263, 131.802, -65.418, -74.887, -69.91]
  MoveL 280 to (-96.75, 392.98, 630.77) mm, rotated rx 170.74 ry 41.15 rz 6.08 deg; joints [-11.098, -30.636, 58.935, 135.123, -69.814, -73.95, -69.91]
  MoveL 281 to (-71.03, 392.99, 602.25) mm, rotated rx 169.88 ry 42.02 rz 6.37 deg; joints [-9.761, -30.824, 60.644, 137.401, -73.478, -72.281, -69.91]
  Set speed (1000.0 mm/s)
  MoveL 282 to (-71.03, 392.99, 602.25) mm, rotated rx 169.88 ry 42.02 rz 6.37 deg; joints [-9.761, -30.824, 60.644, 137.401, -73.478, -72.281, -69.91]
  MoveL 283 to (-7.49, 417.76, 675.38) mm, rotated rx 169.88 ry 42.02 rz 6.37 deg; joints [-6.311, -37.818, 61.155, 140.059, -70.619, -80.01, -69.91]
  Set speed (1000.0 mm/s)
  MoveL 284 to (10.37, 347.65, 672.07) mm, rotated rx 174.15 ry 35.25 rz 4.93 deg; joints [-0.667, -31.666, 55.73, 156.53, -76.5, -89.752, -69.91]
  MoveL 285 to (-45.95, 332.56, 590.83) mm, rotated rx 174.15 ry 35.25 rz 4.93 deg; joints [-4.024, -26.389, 55.997, 151.928, -76.169, -82.858, -69.91]
  MoveL 286 to (-45.95, 332.56, 590.83) mm, rotated rx 174.15 ry 35.25 rz 4.93 deg; joints [-4.024, -26.389, 55.997, 151.928, -76.169, -82.858, -69.91]
  Set speed (50.0 mm/s)
  MoveL 287 to (-72.68, 332.56, 619.57) mm, rotated rx 174.53 ry 35.31 rz 4.6 deg; joints [-5.465, -26.226, 54.702, 149.936, -73.998, -83.815, -69.91]
  MoveL 288 to (-113.93, 332.56, 660.19) mm, rotated rx 174.92 ry 35.36 rz 4.26 deg; joints [-7.761, -25.895, 52.809, 146.266, -70.277, -84.667, -69.91]
  MoveL 289 to (-155.69, 332.56, 700.22) mm, rotated rx 175.3 ry 35.4 rz 3.93 deg; joints [-9.939, -25.384, 50.844, 142.78, -66.75, -85.332, -69.91]
  MoveL 290 to (-198.24, 332.56, 739.35) mm, rotated rx 175.69 ry 35.44 rz 3.6 deg; joints [-12.017, -24.698, 48.812, 139.435, -63.398, -85.815, -69.91]
  MoveL 291 to (-241.81, 332.56, 777.33) mm, rotated rx 176.08 ry 35.48 rz 3.26 deg; joints [-14.009, -23.843, 46.721, 136.2, -60.204, -86.124, -69.91]
  MoveL 292 to (-276.88, 332.56, 806.23) mm, rotated rx 176.47 ry 35.52 rz 2.94 deg; joints [-15.445, -23.002, 45.01, 134.092, -58.087, -86.446, -69.91]
  MoveL 293 to (-312.75, 332.56, 834.2) mm, rotated rx 176.86 ry 35.55 rz 2.61 deg; joints [-16.838, -22.07, 43.267, 132.039, -56.053, -86.692, -69.91]
  MoveL 294 to (-349.49, 332.55, 861.17) mm, rotated rx 176.91 ry 35.56 rz 2.56 deg; joints [-18.473, -21.266, 41.605, 128.504, -52.948, -86.005, -69.91]
  MoveL 295 to (-386.91, 332.55, 886.9) mm, rotated rx 177.28 ry 33.74 rz 2.41 deg; joints [-20.218, -20.232, 39.157, 124.8, -47.376, -86.562, -69.91]
  MoveL 296 to (-425.77, 332.55, 911.82) mm, rotated rx 177.66 ry 31.81 rz 2.22 deg; joints [-21.911, -19.005, 36.566, 121.115, -41.766, -87.03, -69.91]
  MoveL 297 to (-465.33, 332.55, 935.34) mm, rotated rx 178.03 ry 29.82 rz 1.98 deg; joints [-23.524, -17.622, 33.888, 117.438, -36.18, -87.371, -69.91]
  MoveL 298 to (-505.6, 332.55, 957.43) mm, rotated rx 178.41 ry 27.79 rz 1.7 deg; joints [-25.066, -16.097, 31.128, 113.648, -30.545, -87.53, -69.91]
  MoveL 299 to (-546.6, 332.55, 978.06) mm, rotated rx 178.76 ry 25.71 rz 1.39 deg; joints [-26.541, -14.445, 28.285, 109.539, -24.731, -87.402, -69.91]
  MoveL 300 to (-588.35, 332.55, 997.2) mm, rotated rx 179.11 ry 23.61 rz 1.06 deg; joints [-27.957, -12.676, 25.352, 104.68, -18.474, -86.744, -69.91]
  MoveL 301 to (-630.86, 332.55, 1014.83) mm, rotated rx 179.44 ry 21.47 rz 0.7 deg; joints [-29.316, -10.798, 22.289, 97.681, -10.899, -84.747, -69.91]
  MoveL 302 to (-674.14, 332.55, 1030.91) mm, rotated rx 172.93 ry 18.02 rz -20.75 deg; joints [-26.232, -5.473, 17.474, 167.227, -59.713, -109.308, -69.91]
  MoveL 303 to (-718.21, 332.55, 1045.41) mm, rotated rx 174.01 ry 16.08 rz -20.9 deg; joints [-27.528, -3.462, 14.487, 168.551, -57.983, -112.499, -69.91]
  MoveL 304 to (-762.94, 332.55, 1058.27) mm, rotated rx 175.07 ry 14.13 rz -21.08 deg; joints [-28.767, -1.361, 11.437, 170.283, -56.613, -115.792, -69.91]
  MoveL 305 to (-807.9, 332.55, 1069.36) mm, rotated rx 176.07 ry 12.18 rz -21.28 deg; joints [-29.943, 0.805, 8.351, 172.39, -55.608, -119.156, -69.91]
  MoveL 306 to (-853.05, 332.55, 1078.7) mm, rotated rx 177.04 ry 10.23 rz -21.48 deg; joints [-31.061, 3.029, 5.228, 174.838, -54.945, -122.58, -69.91]
  MoveL 307 to (-898.4, 332.55, 1086.31) mm, rotated rx 177.95 ry 8.3 rz -21.68 deg; joints [-32.127, 5.306, 2.065, 177.581, -54.592, -126.049, -69.91]
  MoveL 308 to (-943.92, 332.55, 1092.23) mm, rotated rx 178.82 ry 6.37 rz -21.86 deg; joints [-33.147, 7.633, -1.141, 180.582, -54.518, -129.552, -69.91]
  MoveL 309 to (-989.63, 332.55, 1096.47) mm, rotated rx 179.64 ry 4.45 rz -22.01 deg; joints [-34.127, 10.007, -4.396, 183.801, -54.686, -133.079, -69.91]
  MoveL 310 to (-1031.7, 332.55, 1098.9) mm, rotated rx -179.67 ry 2.69 rz -22.1 deg; joints [-34.995, 12.225, -7.427, 186.908, -55.016, -136.326, -69.91]
  MoveL 311 to (-1073.9, 332.55, 1099.95) mm, rotated rx -179.02 ry 0.93 rz -22.13 deg; joints [-35.838, 14.479, -10.506, 190.133, -55.478, -139.579, -69.91]
  MoveL 312 to (-1116.26, 332.55, 1099.63) mm, rotated rx -178.82 ry -1.31 rz -2.08 deg; joints [-40.186, 13.832, -10.423, 141.445, -4.903, -131.486, -69.91]
  MoveL 313 to (-1158.77, 332.55, 1097.95) mm, rotated rx -178.94 ry -3.14 rz -1.89 deg; joints [-40.714, 16.185, -13.314, 156.402, -11.928, -141.693, -69.91]
  MoveL 314 to (-1201.34, 332.55, 1094.91) mm, rotated rx -179.15 ry -4.95 rz -1.54 deg; joints [-41.306, 18.575, -16.377, 167.271, -16.493, -149.397, -69.91]
  MoveL 315 to (-1243.81, 332.55, 1090.56) mm, rotated rx -179.46 ry -6.72 rz -0.99 deg; joints [-41.926, 20.992, -19.54, 176.741, -20.25, -156.21, -69.91]
  Set speed (1000.0 mm/s)
  MoveL 316 to (-1243.81, 332.55, 1090.56) mm, rotated rx -179.46 ry -6.72 rz -0.99 deg; joints [-41.926, 20.992, -19.54, 176.741, -20.25, -156.21, -69.91]
  MoveL 317 to (-1255.52, 331.81, 1189.87) mm, rotated rx -179.46 ry -6.72 rz -0.99 deg; joints [-41.736, 21.677, -24.077, 191.828, -29.591, -165.884, -69.91]
  Set speed (1000.0 mm/s)
  MoveL 318 to (-1243.18, 271.89, 1190.95) mm, rotated rx -179.84 ry -5.77 rz -0.3 deg; joints [-40.186, 21.8, -24.142, 188.89, -28.587, -163.211, -69.91]
  MoveL 319 to (-1233.12, 272.12, 1091.46) mm, rotated rx -179.84 ry -5.77 rz -0.3 deg; joints [-40.383, 21.206, -19.74, 173.48, -19.208, -153.208, -69.91]
  MoveL 320 to (-1233.12, 272.12, 1091.46) mm, rotated rx -179.84 ry -5.77 rz -0.3 deg; joints [-40.383, 21.206, -19.74, 173.48, -19.208, -153.208, -69.91]
  Set speed (50.0 mm/s)
  MoveL 321 to (-1189.07, 272.12, 1095.24) mm, rotated rx -179.39 ry -4.02 rz -1.09 deg; joints [-39.619, 18.812, -16.577, 165.392, -16.754, -146.961, -69.91]
  MoveL 322 to (-1145.05, 272.12, 1097.65) mm, rotated rx -179.07 ry -2.22 rz -1.65 deg; joints [-38.86, 16.455, -13.495, 157.046, -14.117, -140.553, -69.91]
  MoveL 323 to (-1101.07, 272.12, 1098.68) mm, rotated rx -178.85 ry -0.39 rz -2.01 deg; joints [-38.098, 14.132, -10.493, 148.337, -11.269, -133.9, -69.91]
  MoveL 324 to (-1057.14, 272.12, 1098.31) mm, rotated rx -178.7 ry 1.46 rz -2.21 deg; joints [-37.322, 11.844, -7.572, 139.094, -8.13, -126.888, -69.91]
  MoveL 325 to (-1013.24, 272.13, 1096.51) mm, rotated rx -178.63 ry 3.35 rz -2.29 deg; joints [-36.529, 9.588, -4.741, 128.776, -4.373, -119.193, -69.91]
  MoveL 326 to (-969.39, 272.13, 1093.26) mm, rotated rx 179.5 ry 5.42 rz -22.36 deg; joints [-31.879, 10.529, -4.7, 185.757, -58.613, -131.679, -69.91]
  MoveL 327 to (-921.6, 272.12, 1088.02) mm, rotated rx 178.74 ry 7.39 rz -22.33 deg; joints [-30.752, 8.186, -1.402, 183.099, -59.068, -128.253, -69.91]
  MoveL 328 to (-873.86, 272.12, 1080.98) mm, rotated rx 177.91 ry 9.38 rz -22.25 deg; joints [-29.574, 5.891, 1.857, 180.67, -59.761, -124.853, -69.91]
  MoveL 329 to (-826.46, 272.13, 1072.15) mm, rotated rx -178.84 ry 11.68 rz -1.73 deg; joints [-32.278, 0.358, 7.529, 111.926, -6.068, -101.792, -69.91]
  MoveL 330 to (-779.67, 272.13, 1061.58) mm, rotated rx -179 ry 13.85 rz -1.44 deg; joints [-31.008, -1.846, 10.72, 114.425, -10.862, -101.249, -69.91]
  MoveL 331 to (-733.48, 272.13, 1049.28) mm, rotated rx -179.18 ry 16.02 rz -1.14 deg; joints [-29.693, -3.968, 13.84, 116.5, -15.407, -100.417, -69.91]
  MoveL 332 to (-687.89, 272.12, 1035.27) mm, rotated rx -179.39 ry 18.19 rz -0.81 deg; joints [-28.327, -6.003, 16.901, 118.542, -19.959, -99.513, -69.91]
  MoveL 333 to (-642.89, 272.13, 1019.55) mm, rotated rx -179.62 ry 20.35 rz -0.49 deg; joints [-26.903, -7.946, 19.907, 120.645, -24.583, -98.578, -69.91]
  MoveL 334 to (-598.49, 272.13, 1002.13) mm, rotated rx -179.87 ry 22.5 rz -0.16 deg; joints [-25.417, -9.789, 22.859, 122.854, -29.312, -97.627, -69.91]
  MoveL 335 to (-554.68, 272.13, 983.01) mm, rotated rx 179.86 ry 24.65 rz 0.16 deg; joints [-23.864, -11.522, 25.756, 125.194, -34.167, -96.656, -69.91]
  MoveL 336 to (-511.45, 272.13, 962.2) mm, rotated rx 179.58 ry 26.78 rz 0.46 deg; joints [-22.241, -13.133, 28.595, 127.683, -39.162, -95.658, -69.91]
  MoveL 337 to (-468.82, 272.13, 939.7) mm, rotated rx 179.28 ry 28.88 rz 0.74 deg; joints [-20.542, -14.611, 31.374, 130.337, -44.312, -94.62, -69.91]
  MoveL 338 to (-427.04, 272.13, 915.68) mm, rotated rx 178.97 ry 30.94 rz 1 deg; joints [-18.775, -15.931, 34.069, 133.162, -49.599, -93.539, -69.91]
  MoveL 339 to (-386.35, 272.13, 890.33) mm, rotated rx 178.66 ry 32.95 rz 1.22 deg; joints [-16.949, -17.07, 36.66, 136.163, -55.006, -92.407, -69.91]
  MoveL 340 to (-346.7, 272.13, 863.7) mm, rotated rx 178.35 ry 34.88 rz 1.4 deg; joints [-15.061, -18.017, 39.141, 139.366, -60.55, -91.209, -69.91]
  MoveL 341 to (-308.82, 272.13, 836.43) mm, rotated rx 178.06 ry 36.71 rz 1.54 deg; joints [-13.146, -18.743, 41.46, 142.734, -66.134, -89.957, -69.91]
  MoveL 342 to (-271.86, 272.13, 808.04) mm, rotated rx 177.78 ry 38.46 rz 1.63 deg; joints [-11.165, -19.251, 43.657, 146.371, -71.893, -88.613, -69.91]
  MoveL 343 to (-235.78, 272.13, 778.58) mm, rotated rx -166.07 ry 38.07 rz 27.4 deg; joints [-14.902, -23.833, 47.176, 100.01, -42.034, -80.435, -69.91]
  MoveL 344 to (-200.52, 272.13, 748.11) mm, rotated rx -165.35 ry 39.53 rz 27.96 deg; joints [-12.857, -24.104, 49.361, 107.239, -49.363, -82.607, -69.91]
  MoveL 345 to (-156.75, 272.13, 708) mm, rotated rx -164.95 ry 39.69 rz 27.83 deg; joints [-10.143, -24.159, 51.31, 115.085, -55.603, -85.355, -69.91]
  MoveL 346 to (-114.09, 272.13, 666.52) mm, rotated rx -164.43 ry 40.61 rz 28.18 deg; joints [-7.402, -23.949, 53.462, 122.384, -62.92, -86.616, -69.91]
  MoveL 347 to (-72.38, 272.13, 623.9) mm, rotated rx -163.89 ry 41.52 rz 28.54 deg; joints [-4.535, -23.364, 55.462, 129.581, -70.434, -87.173, -69.91]
  MoveL 348 to (-31.38, 272.13, 580.41) mm, rotated rx -148.72 ry 34.17 rz 52.25 deg; joints [-8.292, -27.899, 57.713, 81.467, -39.389, -78.296, -69.91]
  Set speed (1000.0 mm/s)
  MoveL 349 to (-31.38, 272.13, 580.41) mm, rotated rx -148.72 ry 34.17 rz 52.25 deg; joints [-8.292, -27.899, 57.713, 81.467, -39.389, -78.296, -69.91]
  MoveL 350 to (39.06, 278.29, 651.12) mm, rotated rx -148.72 ry 34.17 rz 52.25 deg; joints [-3.844, -33.437, 57.762, 82.442, -33.147, -83.972, -69.91]
  Set speed (1000.0 mm/s)
  MoveL 351 to (54.39, 213.78, 636.81) mm, rotated rx -144.33 ry 35.57 rz 52.56 deg; joints [1.643, -26.878, 56.731, 107.541, -53.282, -96.48, -69.91]
  MoveL 352 to (-20.64, 211.7, 570.73) mm, rotated rx -144.33 ry 35.57 rz 52.56 deg; joints [-3.194, -22.027, 56.542, 103.424, -56.288, -89.719, -69.91]
  MoveL 353 to (-20.64, 211.7, 570.73) mm, rotated rx -144.33 ry 35.57 rz 52.56 deg; joints [-3.194, -22.027, 56.542, 103.424, -56.288, -89.719, -69.91]
  Set speed (50.0 mm/s)
  MoveL 354 to (-52.78, 211.7, 606.53) mm, rotated rx -145.59 ry 35.12 rz 52.35 deg; joints [-5.763, -23.22, 55.075, 94.146, -48.626, -86.097, -69.91]
  MoveL 355 to (-85.54, 211.7, 641.56) mm, rotated rx -146.88 ry 34.44 rz 51.9 deg; joints [-8.109, -24.017, 53.335, 84.292, -40.617, -81.708, -69.91]
  MoveL 356 to (-119.01, 211.7, 675.73) mm, rotated rx -148.19 ry 33.59 rz 51.29 deg; joints [-10.227, -24.452, 51.356, 73.126, -31.913, -76.124, -69.91]
  MoveL 357 to (-153.25, 211.7, 708.96) mm, rotated rx -163.34 ry 40.72 rz 27.67 deg; joints [-6.764, -20.295, 49.51, 125.202, -64.545, -88.997, -69.91]
  MoveL 358 to (-188.29, 211.7, 741.2) mm, rotated rx -164.14 ry 39.26 rz 27.05 deg; joints [-8.944, -20.509, 47.559, 119.31, -57.52, -88.498, -69.91]
  MoveL 359 to (-223.53, 211.7, 771.84) mm, rotated rx -164.9 ry 37.73 rz 26.41 deg; joints [-11.008, -20.443, 45.489, 113.388, -50.582, -87.607, -69.91]
  MoveL 360 to (-259.63, 211.7, 801.43) mm, rotated rx -165.63 ry 36.11 rz 25.75 deg; joints [-12.997, -20.127, 43.275, 107.099, -43.483, -86.217, -69.91]
  MoveL 361 to (-296.63, 211.7, 829.92) mm, rotated rx 179.27 ry 36.72 rz 0.58 deg; joints [-9.768, -15.527, 39.442, 151.833, -73.974, -92.539, -69.91]
  MoveL 362 to (-334.55, 211.7, 857.27) mm, rotated rx 179.5 ry 34.89 rz 0.42 deg; joints [-11.699, -14.982, 37.231, 148.728, -68.5, -94.208, -69.91]
  MoveL 363 to (-374.24, 211.7, 883.96) mm, rotated rx 179.75 ry 32.96 rz 0.23 deg; joints [-13.621, -14.22, 34.864, 145.839, -63.104, -95.816, -69.91]
  MoveL 364 to (-414.96, 211.7, 909.37) mm, rotated rx 179.99 ry 30.98 rz 0.01 deg; joints [-15.493, -13.262, 32.39, 143.21, -57.89, -97.355, -69.91]
  MoveL 365 to (-456.76, 211.7, 933.47) mm, rotated rx -179.77 ry 28.95 rz -0.24 deg; joints [-17.316, -12.123, 29.814, 140.831, -52.849, -98.856, -69.91]
  MoveL 366 to (-499.64, 211.7, 956.18) mm, rotated rx -179.54 ry 26.87 rz -0.5 deg; joints [-19.088, -10.812, 27.141, 138.701, -47.982, -100.344, -69.91]
  MoveL 367 to (-543.2, 211.7, 977.25) mm, rotated rx -179.32 ry 24.78 rz -0.78 deg; joints [-20.792, -9.356, 24.4, 136.844, -43.337, -101.836, -69.91]
  MoveL 368 to (-587.31, 211.7, 996.62) mm, rotated rx -179.12 ry 22.67 rz -1.07 deg; joints [-22.426, -7.771, 21.604, 135.282, -38.935, -103.36, -69.91]
  MoveL 369 to (-631.97, 211.7, 1014.29) mm, rotated rx -178.93 ry 20.56 rz -1.36 deg; joints [-23.991, -6.07, 18.757, 134.038, -34.791, -104.952, -69.91]
  MoveL 370 to (-677.17, 211.7, 1030.26) mm, rotated rx -178.76 ry 18.44 rz -1.65 deg; joints [-25.49, -4.264, 15.862, 133.149, -30.922, -106.651, -69.91]
  MoveL 371 to (-722.91, 211.7, 1044.54) mm, rotated rx -178.61 ry 16.33 rz -1.92 deg; joints [-26.926, -2.361, 12.922, 132.673, -27.361, -108.507, -69.91]
  MoveL 372 to (-769.2, 211.7, 1057.13) mm, rotated rx -178.49 ry 14.22 rz -2.17 deg; joints [-28.302, -0.369, 9.938, 132.698, -24.159, -110.586, -69.91]
  MoveL 373 to (-816.03, 211.7, 1068.02) mm, rotated rx -178.39 ry 12.11 rz -2.39 deg; joints [-29.62, 1.707, 6.911, 133.336, -21.381, -112.962, -69.91]
  MoveL 374 to (-863.4, 211.7, 1077.21) mm, rotated rx -178.33 ry 10.01 rz -2.56 deg; joints [-30.882, 3.86, 3.843, 134.716, -19.105, -115.722, -69.91]
  MoveL 375 to (-911.32, 211.7, 1084.7) mm, rotated rx -178.32 ry 7.93 rz -2.66 deg; joints [-32.09, 6.087, 0.733, 136.987, -17.419, -118.96, -69.91]
  MoveL 376 to (-959.49, 211.7, 1090.45) mm, rotated rx -178.35 ry 5.86 rz -2.68 deg; joints [-33.24, 8.371, -2.401, 140.24, -16.392, -122.727, -69.91]
  MoveL 377 to (-1003.68, 211.7, 1094.2) mm, rotated rx -178.43 ry 4 rz -2.6 deg; joints [-34.242, 10.503, -5.29, 144.078, -16.028, -126.64, -69.91]
  MoveL 378 to (-1047.91, 211.7, 1096.53) mm, rotated rx -178.58 ry 2.17 rz -2.41 deg; joints [-35.202, 12.67, -8.202, 148.639, -16.145, -130.946, -69.91]
  MoveL 379 to (-1092.17, 211.7, 1097.46) mm, rotated rx -178.8 ry 0.36 rz -2.08 deg; joints [-36.128, 14.87, -11.146, 153.797, -16.647, -135.581, -69.91]
  MoveL 380 to (-1136.47, 211.7, 1097.03) mm, rotated rx -179.1 ry -1.41 rz -1.58 deg; joints [-37.027, 17.103, -14.132, 159.41, -17.422, -140.473, -69.91]
  MoveL 381 to (-1180.81, 211.7, 1095.26) mm, rotated rx -179.51 ry -3.14 rz -0.87 deg; joints [-37.911, 19.371, -17.167, 165.363, -18.366, -145.575, -69.91]
  MoveL 382 to (-1225.17, 211.7, 1092.16) mm, rotated rx 179.95 ry -4.83 rz 0.09 deg; joints [-38.788, 21.674, -20.258, 171.594, -19.403, -150.87, -69.91]
  Set speed (1000.0 mm/s)
  MoveL 383 to (-1225.17, 211.7, 1092.16) mm, rotated rx 179.95 ry -4.83 rz 0.09 deg; joints [-38.788, 21.674, -20.258, 171.594, -19.403, -150.87, -69.91]
  MoveL 384 to (-1233.59, 211.77, 1191.81) mm, rotated rx 179.95 ry -4.83 rz 0.09 deg; joints [-38.593, 22.188, -24.55, 186.686, -28.467, -160.795, -69.91]
  Set speed (1000.0 mm/s)
  MoveL 385 to (-1226.38, 151.48, 1192.45) mm, rotated rx 179.86 ry -3.87 rz 0.24 deg; joints [-36.977, 22.816, -25.265, 185.218, -29.115, -158.709, -69.91]
  MoveL 386 to (-1219.62, 151.27, 1092.68) mm, rotated rx 179.86 ry -3.87 rz 0.24 deg; joints [-37.166, 22.371, -21.063, 170.94, -20.626, -149.181, -69.91]
  MoveL 387 to (-1219.62, 151.27, 1092.68) mm, rotated rx 179.86 ry -3.87 rz 0.24 deg; joints [-37.166, 22.371, -21.063, 170.94, -20.626, -149.181, -69.91]
  Set speed (50.0 mm/s)
  MoveL 388 to (-1175.09, 151.27, 1095.07) mm, rotated rx -179.53 ry -2.26 rz -0.83 deg; joints [-36.198, 20.161, -18.039, 166.356, -20.785, -144.767, -69.91]
  MoveL 389 to (-1130.61, 151.27, 1096.2) mm, rotated rx -179.05 ry -0.6 rz -1.65 deg; joints [-35.222, 17.988, -15.059, 162.125, -21.042, -140.612, -69.91]
  MoveL 390 to (-1086.19, 151.27, 1096.04) mm, rotated rx -178.69 ry 1.1 rz -2.25 deg; joints [-34.231, 15.849, -12.12, 158.246, -21.437, -136.693, -69.91]
  MoveL 391 to (-1041.84, 151.27, 1094.57) mm, rotated rx -178.41 ry 2.84 rz -2.68 deg; joints [-33.217, 13.745, -9.215, 154.743, -22.022, -133.006, -69.91]
  MoveL 392 to (-997.55, 151.27, 1091.76) mm, rotated rx -178.21 ry 4.61 rz -2.95 deg; joints [-32.175, 11.676, -6.341, 151.65, -22.843, -129.552, -69.91]
  MoveL 393 to (-953.32, 151.27, 1087.58) mm, rotated rx -178.07 ry 6.41 rz -3.11 deg; joints [-31.098, 9.644, -3.491, 148.992, -23.942, -126.332, -69.91]
  MoveL 394 to (-905.15, 151.27, 1081.42) mm, rotated rx -177.98 ry 8.41 rz -3.17 deg; joints [-29.876, 7.473, -0.409, 146.62, -25.496, -123.09, -69.91]
  MoveL 395 to (-857.09, 151.27, 1073.55) mm, rotated rx -177.94 ry 10.44 rz -3.13 deg; joints [-28.6, 5.354, 2.65, 144.807, -27.443, -120.123, -69.91]
  MoveL 396 to (-809.48, 151.27, 1064.01) mm, rotated rx -177.95 ry 12.48 rz -3.02 deg; joints [-27.273, 3.307, 5.664, 143.548, -29.77, -117.429, -69.91]
  MoveL 397 to (-762.46, 151.27, 1052.81) mm, rotated rx -178 ry 14.54 rz -2.86 deg; joints [-25.896, 1.343, 8.628, 142.806, -32.457, -114.979, -69.91]
  MoveL 398 to (-716.02, 151.27, 1039.98) mm, rotated rx -178.07 ry 16.6 rz -2.65 deg; joints [-24.465, -0.532, 11.541, 142.539, -35.484, -112.737, -69.91]
  MoveL 399 to (-670.15, 151.27, 1025.49) mm, rotated rx -178.17 ry 18.66 rz -2.42 deg; joints [-22.977, -2.312, 14.404, 142.704, -38.829, -110.666, -69.91]
  MoveL 400 to (-624.87, 151.27, 1009.35) mm, rotated rx -178.29 ry 20.73 rz -2.16 deg; joints [-21.43, -3.99, 17.214, 143.257, -42.468, -108.726, -69.91]
  MoveL 401 to (-580.18, 151.27, 991.57) mm, rotated rx -178.43 ry 22.8 rz -1.9 deg; joints [-19.823, -5.555, 19.972, 144.165, -46.385, -106.881, -69.91]
  MoveL 402 to (-536.06, 151.27, 972.14) mm, rotated rx -178.58 ry 24.86 rz -1.63 deg; joints [-18.153, -6.999, 22.673, 145.404, -50.57, -105.097, -69.91]
  MoveL 403 to (-492.53, 151.27, 951.05) mm, rotated rx -178.75 ry 26.91 rz -1.37 deg; joints [-16.42, -8.308, 25.314, 146.958, -55.01, -103.344, -69.91]
  MoveL 404 to (-449.57, 151.27, 928.3) mm, rotated rx -178.93 ry 28.96 rz -1.11 deg; joints [-14.623, -9.471, 27.891, 148.818, -59.702, -101.587, -69.91]
  MoveL 405 to (-407.43, 151.27, 904.02) mm, rotated rx -179.11 ry 30.97 rz -0.86 deg; joints [-12.771, -10.468, 30.387, 150.972, -64.622, -99.805, -69.91]
  MoveL 406 to (-366.38, 151.27, 878.42) mm, rotated rx -179.3 ry 32.95 rz -0.64 deg; joints [-10.881, -11.279, 32.777, 153.406, -69.734, -97.978, -69.91]
  MoveL 407 to (-326.4, 151.27, 851.56) mm, rotated rx -179.49 ry 34.87 rz -0.43 deg; joints [-8.952, -11.894, 35.059, 156.128, -75.041, -96.074, -69.91]
  MoveL 408 to (-288.22, 151.27, 824.03) mm, rotated rx -165.41 ry 34.07 rz 24.14 deg; joints [-11.733, -16.485, 39.154, 112.633, -44.009, -90.963, -69.91]
  MoveL 409 to (-251, 151.27, 795.36) mm, rotated rx -164.67 ry 35.76 rz 24.83 deg; joints [-9.782, -16.863, 41.382, 118.207, -50.823, -91.861, -69.91]
  MoveL 410 to (-214.72, 151.28, 765.58) mm, rotated rx -163.9 ry 37.39 rz 25.53 deg; joints [-7.787, -17.015, 43.484, 123.451, -57.497, -92.303, -69.91]
  MoveL 411 to (-179.33, 151.28, 734.73) mm, rotated rx -163.12 ry 38.97 rz 26.24 deg; joints [-5.75, -16.924, 45.455, 128.552, -64.138, -92.359, -69.91]
  MoveL 412 to (-144.2, 151.28, 702.25) mm, rotated rx -162.29 ry 40.5 rz 26.94 deg; joints [-3.633, -16.562, 47.32, 133.74, -70.943, -92.059, -69.91]
  MoveL 413 to (-109.94, 151.28, 668.73) mm, rotated rx -147.38 ry 33.18 rz 50.43 deg; joints [-6.926, -20.724, 49.604, 86.854, -39.397, -84.459, -69.91]
  MoveL 414 to (-76.53, 151.28, 634.2) mm, rotated rx -146 ry 34.19 rz 51.25 deg; joints [-4.823, -20.112, 51.506, 95.937, -47.607, -88.087, -69.91]
  MoveL 415 to (-43.92, 151.28, 598.71) mm, rotated rx -144.62 ry 35.09 rz 52 deg; joints [-2.607, -19.159, 53.208, 104.167, -55.458, -90.764, -69.91]
  MoveL 416 to (-12.09, 151.28, 562.31) mm, rotated rx -143.25 ry 35.87 rz 52.65 deg; joints [-0.281, -17.84, 54.693, 111.987, -63.153, -92.728, -69.91]
  Set speed (1000.0 mm/s)
  MoveL 417 to (-12.09, 151.28, 562.31) mm, rotated rx -143.25 ry 35.87 rz 52.65 deg; joints [-0.281, -17.84, 54.693, 111.987, -63.153, -92.728, -69.91]
  MoveL 418 to (63.96, 152.3, 627.24) mm, rotated rx -143.25 ry 35.87 rz 52.65 deg; joints [4.465, -22.281, 54.878, 116.331, -60.997, -99.112, -69.91]
  Set speed (1000.0 mm/s)
  MoveL 419 to (70.5, 91.94, 619.89) mm, rotated rx -143.14 ry 35.96 rz 52.75 deg; joints [6.281, -18.528, 52.865, 120.979, -65.204, -99.704, -69.91]
  MoveL 420 to (-5.68, 90.85, 555.13) mm, rotated rx -143.14 ry 35.96 rz 52.75 deg; joints [1.739, -14.353, 52.68, 116.784, -67.007, -93.732, -69.91]
  MoveL 421 to (-5.68, 90.85, 555.13) mm, rotated rx -143.14 ry 35.96 rz 52.75 deg; joints [1.739, -14.353, 52.68, 116.784, -67.007, -93.732, -69.91]
  Set speed (50.0 mm/s)
  MoveL 422 to (-37.49, 90.85, 591.87) mm, rotated rx -144.62 ry 35.09 rz 52 deg; joints [-0.507, -15.791, 51.264, 109.414, -59.3, -92.337, -69.91]
  MoveL 423 to (-70.13, 90.85, 627.64) mm, rotated rx -146.1 ry 34.15 rz 51.24 deg; joints [-2.712, -16.898, 49.663, 101.582, -51.479, -90.15, -69.91]
  MoveL 424 to (-103.63, 90.85, 662.4) mm, rotated rx -147.59 ry 33.15 rz 50.48 deg; joints [-4.861, -17.69, 47.884, 92.927, -43.37, -86.984, -69.91]
  MoveL 425 to (-138.02, 90.85, 696.12) mm, rotated rx -149.07 ry 32.1 rz 49.72 deg; joints [-6.931, -18.185, 45.923, 82.821, -34.638, -82.474, -69.91]
  MoveL 426 to (-173.31, 90.85, 728.77) mm, rotated rx -163.59 ry 38.9 rz 26.46 deg; joints [-4.011, -14.332, 43.733, 131.397, -66.517, -92.389, -69.91]
  MoveL 427 to (-208.88, 90.85, 759.77) mm, rotated rx -164.52 ry 37.36 rz 25.91 deg; joints [-6.119, -14.619, 41.896, 125.896, -59.592, -92.194, -69.91]
  MoveL 428 to (-245.37, 90.85, 789.68) mm, rotated rx -165.44 ry 35.78 rz 25.38 deg; joints [-8.205, -14.667, 39.926, 120.134, -52.572, -91.511, -69.91]
  MoveL 429 to (-282.81, 90.85, 818.48) mm, rotated rx -166.33 ry 34.14 rz 24.87 deg; joints [-10.262, -14.487, 37.822, 113.886, -45.332, -90.242, -69.91]
  MoveL 430 to (-321.22, 90.84, 846.13) mm, rotated rx 179.44 ry 34.63 rz 0.48 deg; joints [-7.72, -10.2, 33.756, 155.989, -74.904, -94.826, -69.91]
  MoveL 431 to (-361.46, 90.85, 873.12) mm, rotated rx 179.46 ry 32.71 rz 0.49 deg; joints [-9.745, -9.782, 31.613, 152.527, -68.977, -96.432, -69.91]
  MoveL 432 to (-402.77, 90.85, 898.85) mm, rotated rx 179.49 ry 30.75 rz 0.5 deg; joints [-11.742, -9.16, 29.354, 149.249, -63.173, -97.884, -69.91]
  MoveL 433 to (-445.15, 90.85, 923.23) mm, rotated rx 179.51 ry 28.76 rz 0.51 deg; joints [-13.704, -8.344, 26.984, 146.134, -57.485, -99.204, -69.91]
  MoveL 434 to (-488.17, 90.85, 946) mm, rotated rx 179.54 ry 26.75 rz 0.51 deg; joints [-15.607, -7.353, 24.531, 143.186, -51.961, -100.398, -69.91]
  MoveL 435 to (-531.75, 90.85, 967.12) mm, rotated rx 179.56 ry 24.75 rz 0.51 deg; joints [-17.444, -6.202, 22.004, 140.392, -46.601, -101.489, -69.91]
  MoveL 436 to (-575.88, 90.85, 986.6) mm, rotated rx 179.58 ry 22.73 rz 0.51 deg; joints [-19.213, -4.904, 19.405, 137.736, -41.393, -102.496, -69.91]
  MoveL 437 to (-620.55, 90.85, 1004.45) mm, rotated rx 179.6 ry 20.73 rz 0.5 deg; joints [-20.911, -3.47, 16.739, 135.208, -36.337, -103.437, -69.91]
  MoveL 438 to (-665.76, 90.85, 1020.68) mm, rotated rx 179.63 ry 18.74 rz 0.49 deg; joints [-22.539, -1.909, 14.005, 132.803, -31.432, -104.329, -69.91]
  MoveL 439 to (-711.52, 90.84, 1035.29) mm, rotated rx 179.65 ry 16.76 rz 0.48 deg; joints [-24.096, -0.231, 11.205, 130.529, -26.678, -105.197, -69.91]
  MoveL 440 to (-757.81, 90.84, 1048.3) mm, rotated rx 179.67 ry 14.79 rz 0.47 deg; joints [-25.582, 1.557, 8.337, 128.413, -22.088, -106.073, -69.91]
  MoveL 441 to (-804.63, 90.84, 1059.7) mm, rotated rx 179.69 ry 12.85 rz 0.45 deg; joints [-26.997, 3.45, 5.404, 126.507, -17.701, -106.999, -69.91]
  MoveL 442 to (-851.99, 90.84, 1069.51) mm, rotated rx 179.71 ry 10.93 rz 0.43 deg; joints [-28.34, 5.442, 2.403, 124.953, -13.603, -108.072, -69.91]
  MoveL 443 to (-899.88, 90.84, 1077.74) mm, rotated rx 179.74 ry 9.04 rz 0.41 deg; joints [-29.608, 7.53, -0.659, 124.112, -10.017, -109.513, -69.91]
  MoveL 444 to (-948.28, 90.84, 1084.38) mm, rotated rx 179.76 ry 7.18 rz 0.38 deg; joints [-30.792, 9.711, -3.766, 124.92, -7.54, -111.878, -69.91]
  MoveL 445 to (-1001.72, 90.84, 1089.82) mm, rotated rx 179.79 ry 5.18 rz 0.34 deg; joints [-31.961, 12.198, -7.177, 129.583, -7.315, -116.628, -69.91]
  MoveL 446 to (-1055.24, 90.84, 1093.34) mm, rotated rx 179.82 ry 3.25 rz 0.3 deg; joints [-32.984, 14.77, -10.605, 138.043, -9.66, -123.511, -69.91]
  MoveL 447 to (-1108.82, 90.84, 1095.02) mm, rotated rx 179.86 ry 1.37 rz 0.24 deg; joints [-33.892, 17.43, -14.136, 148.028, -13.204, -131.153, -69.91]
  MoveL 448 to (-1162.47, 90.84, 1094.9) mm, rotated rx 179.9 ry -0.44 rz 0.17 deg; joints [-34.716, 20.182, -17.825, 158.25, -17.202, -138.753, -69.91]
  MoveL 449 to (-1216.18, 90.84, 1093.02) mm, rotated rx 179.94 ry -2.17 rz 0.11 deg; joints [-35.485, 23.018, -21.682, 167.982, -21.236, -145.857, -69.91]
  Set speed (1000.0 mm/s)
  MoveL 450 to (-1216.18, 90.84, 1093.02) mm, rotated rx 179.94 ry -2.17 rz 0.11 deg; joints [-35.485, 23.018, -21.682, 167.982, -21.236, -145.857, -69.91]
  MoveL 451 to (-1219.97, 90.95, 1192.95) mm, rotated rx 179.94 ry -2.17 rz 0.11 deg; joints [-35.273, 23.331, -25.696, 181.575, -29.139, -155.132, -69.91]
  Set speed (1000.0 mm/s)
  MoveL 452 to (-1217.51, 30.46, 1193.15) mm, rotated rx 179.97 ry -1.68 rz 0.05 deg; joints [-33.712, 24.599, -27.338, 183.242, -31.788, -154.934, -69.91]
  MoveL 453 to (-1214.58, 30.42, 1093.19) mm, rotated rx 179.97 ry -1.68 rz 0.05 deg; joints [-33.902, 24.288, -23.3, 171.097, -24.698, -146.536, -69.91]
  MoveL 454 to (-1214.58, 30.42, 1093.19) mm, rotated rx 179.97 ry -1.68 rz 0.05 deg; joints [-33.902, 24.288, -23.3, 171.097, -24.698, -146.536, -69.91]
  Set speed (50.0 mm/s)
  MoveL 455 to (-1160.74, 30.42, 1094.2) mm, rotated rx 179.96 ry 0.02 rz 0.07 deg; joints [-33.062, 21.479, -19.373, 162.836, -21.595, -140.289, -69.91]
  MoveL 456 to (-1106.98, 30.42, 1093.54) mm, rotated rx 179.95 ry 1.79 rz 0.09 deg; joints [-32.153, 18.777, -15.622, 154.963, -19.048, -134.084, -69.91]
  MoveL 457 to (-1053.31, 30.42, 1091.18) mm, rotated rx 179.94 ry 3.62 rz 0.11 deg; joints [-31.156, 16.173, -12.014, 147.973, -17.327, -128.237, -69.91]
  MoveL 458 to (-999.72, 30.42, 1087.05) mm, rotated rx 179.93 ry 5.52 rz 0.12 deg; joints [-30.058, 13.662, -8.508, 142.402, -16.728, -123.091, -69.91]
  MoveL 459 to (-946.22, 30.42, 1081.08) mm, rotated rx 179.92 ry 7.47 rz 0.13 deg; joints [-28.848, 11.243, -5.074, 138.608, -17.436, -118.878, -69.91]
  MoveL 460 to (-897.79, 30.42, 1074.04) mm, rotated rx 179.91 ry 9.3 rz 0.14 deg; joints [-27.652, 9.129, -2.003, 136.68, -19.17, -115.859, -69.91]
  MoveL 461 to (-849.84, 30.42, 1065.46) mm, rotated rx 179.9 ry 11.17 rz 0.14 deg; joints [-26.376, 7.111, 1.004, 135.94, -21.743, -113.475, -69.91]
  MoveL 462 to (-802.42, 30.42, 1055.35) mm, rotated rx 179.9 ry 13.06 rz 0.15 deg; joints [-25.024, 5.193, 3.946, 136.075, -24.947, -111.541, -69.91]
  MoveL 463 to (-755.52, 30.42, 1043.68) mm, rotated rx 179.89 ry 14.98 rz 0.15 deg; joints [-23.599, 3.378, 6.823, 136.832, -28.62, -109.9, -69.91]
  MoveL 464 to (-709.15, 30.42, 1030.46) mm, rotated rx 179.89 ry 16.93 rz 0.16 deg; joints [-22.103, 1.67, 9.637, 138.039, -32.653, -108.439, -69.91]
  MoveL 465 to (-663.31, 30.42, 1015.66) mm, rotated rx 179.88 ry 18.89 rz 0.16 deg; joints [-20.538, 0.078, 12.382, 139.59, -36.972, -107.089, -69.91]
  MoveL 466 to (-618.01, 30.42, 999.28) mm, rotated rx 179.87 ry 20.87 rz 0.16 deg; joints [-18.906, -1.393, 15.06, 141.416, -41.532, -105.791, -69.91]
  MoveL 467 to (-573.24, 30.42, 981.31) mm, rotated rx 179.87 ry 22.86 rz 0.16 deg; joints [-17.206, -2.733, 17.67, 143.474, -46.312, -104.501, -69.91]
  MoveL 468 to (-529.02, 30.42, 961.73) mm, rotated rx 179.86 ry 24.86 rz 0.16 deg; joints [-15.443, -3.934, 20.21, 145.745, -51.295, -103.186, -69.91]
  MoveL 469 to (-485.35, 30.42, 940.54) mm, rotated rx 179.85 ry 26.86 rz 0.16 deg; joints [-13.618, -4.985, 22.675, 148.222, -56.467, -101.821, -69.91]
  MoveL 470 to (-442.22, 30.42, 917.71) mm, rotated rx 179.85 ry 28.86 rz 0.16 deg; joints [-11.734, -5.873, 25.063, 150.907, -61.831, -100.375, -69.91]
  MoveL 471 to (-399.75, 30.42, 893.28) mm, rotated rx 179.84 ry 30.85 rz 0.16 deg; joints [-9.8, -6.585, 27.366, 153.804, -67.381, -98.822, -69.91]
  MoveL 472 to (-358.32, 30.42, 867.53) mm, rotated rx 179.83 ry 32.8 rz 0.15 deg; joints [-7.838, -7.105, 29.555, 156.903, -73.063, -97.154, -69.91]
  MoveL 473 to (-317.97, 30.42, 840.5) mm, rotated rx -166.82 ry 32.41 rz 24.05 deg; joints [-10.107, -11.355, 33.779, 114.395, -42.936, -91.815, -69.91]
  MoveL 474 to (-279.44, 30.42, 812.82) mm, rotated rx -165.93 ry 34.08 rz 24.53 deg; joints [-8.112, -11.637, 35.918, 120.475, -50.091, -93.07, -69.91]
  MoveL 475 to (-241.88, 30.42, 783.99) mm, rotated rx -165.03 ry 35.71 rz 25.05 deg; joints [-6.095, -11.708, 37.926, 126.016, -56.98, -93.743, -69.91]
  MoveL 476 to (-205.27, 30.42, 754.05) mm, rotated rx -164.11 ry 37.29 rz 25.59 deg; joints [-4.064, -11.56, 39.805, 131.247, -63.727, -93.946, -69.91]
  MoveL 477 to (-169.59, 30.42, 723.02) mm, rotated rx -163.17 ry 38.83 rz 26.16 deg; joints [-2.024, -11.184, 41.554, 136.324, -70.42, -93.737, -69.91]
  MoveL 478 to (-134.17, 30.42, 690.34) mm, rotated rx -148.76 ry 31.91 rz 49.33 deg; joints [-4.764, -14.963, 43.996, 91.128, -39.534, -86.978, -69.91]
  MoveL 479 to (-99.67, 30.42, 656.58) mm, rotated rx -147.28 ry 32.97 rz 50.11 deg; joints [-2.72, -14.369, 45.842, 99.874, -47.676, -90.372, -69.91]
  MoveL 480 to (-66.05, 30.42, 621.79) mm, rotated rx -145.81 ry 33.98 rz 50.91 deg; joints [-0.636, -13.499, 47.519, 107.562, -55.376, -92.699, -69.91]
  MoveL 481 to (-33.29, 30.42, 585.97) mm, rotated rx -144.35 ry 34.94 rz 51.71 deg; joints [1.472, -12.343, 49.031, 114.624, -62.861, -94.202, -69.91]
  MoveL 482 to (-1.38, 30.42, 549.16) mm, rotated rx -142.89 ry 35.85 rz 52.53 deg; joints [3.594, -10.89, 50.374, 121.328, -70.258, -95.011, -69.91]
  Set speed (1000.0 mm/s)
  MoveL 483 to (-1.38, 30.42, 549.16) mm, rotated rx -142.89 ry 35.85 rz 52.53 deg; joints [3.594, -10.89, 50.374, 121.328, -70.258, -95.011, -69.91]
  MoveL 484 to (74.91, 30.79, 613.8) mm, rotated rx -142.89 ry 35.85 rz 52.53 deg; joints [7.934, -14.76, 50.523, 125.444, -68.849, -100.596, -69.91]

